Omron Sysmac Studio project 3089-2603A_検査箱詰め装置_CORE_SUB_PIP-02F02NX_20261026D (Sysmac Studio 1.67.0.7, StandardProject)
(* イーサキャット設定完了_20261023I / ST0 供給_20261009A / AutoMode作成_20261008A / IOプログラム作成_20261007B / IOプログラム作成_20261006A / IOプログラム作成_20261005A / IOプログラム作成_20261002A / オリエンタルモータ設定_20261001A / IO設定_20260930A / PLC設定_20260807A *)

# Controller new_Controller_0: NX102-9020 version 1.48
Units and slaves: Node1 : RCGW-ECT(112Byte/112Byte) (E001); Node2 : CVD2A-KED (E002); Node3 : CVD2A-KED (E003); Node5 : RCGW-ECT(112Byte/112Byte) (E005); Node6 : GX-ID1612 (E006); Node7 : GX-ID1612 (E007); Node8 : GX-OD1612 (E008); Node9 : GX-ID1612 (E011); Node10 : GX-OD1612 (E010); ユニット1 : NX-ID6142-6(N1); ユニット2 : NX-ID6142-6(N2); ユニット3 : NX-ID6142-6(N3); ユニット4 : NX-ID6142-6(N4); ユニット5 : NX-ID6142-6(N5); ユニット6 : NX-OD6121-6(N6); ユニット7 : NX-OD6121-6(N7); ユニット8 : NX-OD6121-6(N8)
Axis Stm_A_Rev_Axis000, settings changed from default: AxisType=ServoType, FunctionLimit=SingleAxisPTP, UnitsConversion=EnumElement5, UnitsDenominator=360, MaxVelocity=10000, MaxJogVelocity=10000, HomingMode=BackupAndProximitySignalOn, OriginInputMode=EXT, StartDirection=NegativeDirection, OriginInputDetectionDirection=NegativeDirection, CountMode=EnumElement2, ModuloMAXPosition=360, ModuloMINPosition=0
Axis Stm_A_Rev_Axis001, settings changed from default: AxisNumber=1, AxisType=ServoType, FunctionLimit=SingleAxisPTP, UnitsConversion=EnumElement5, UnitsDenominator=360, MaxVelocity=10000, MaxJogVelocity=10000, HomingMode=BackupAndProximitySignalOn, OriginInputMode=EXT, StartDirection=NegativeDirection, OriginInputDetectionDirection=NegativeDirection, CountMode=EnumElement2, ModuloMAXPosition=360, ModuloMINPosition=0
Axis Stm_B_Rev_Axis002, settings changed from default: AxisNumber=2, AxisType=ServoType, FunctionLimit=SingleAxisPTP, UnitsConversion=EnumElement5, UnitsDenominator=360, MaxVelocity=10000, MaxJogVelocity=10000, HomingMode=BackupAndProximitySignalOn, OriginInputMode=EXT, StartDirection=NegativeDirection, OriginInputDetectionDirection=NegativeDirection, CountMode=EnumElement2, ModuloMAXPosition=360, ModuloMINPosition=0
Axis Stm_B_Rev_Axis003, settings changed from default: AxisNumber=3, AxisType=ServoType, FunctionLimit=SingleAxisPTP, UnitsConversion=EnumElement5, UnitsDenominator=360, MaxVelocity=10000, MaxJogVelocity=10000, HomingMode=BackupAndProximitySignalOn, OriginInputMode=EXT, StartDirection=NegativeDirection, OriginInputDetectionDirection=NegativeDirection, CountMode=EnumElement2, ModuloMAXPosition=360, ModuloMINPosition=0
Task PrimaryTask (priority 4, period or condition 2000): ModeManagement_モード管理, Movements_動作, OtherDevice_外部機器, IO_入出力

TYPE sData : STRUCT
    Dates : STRING[20];  (* 検査日時 *)
    Work_On : BOOL;  (* ワーク有無(0:無 1:有) *)
    Total_Judge : INT;  (* 総合判定(0:無 1:OK 9:NG) *)
    Judgment_Details : INT;  (* NG内容 *)
    HeightData : LREAL;  (* 高さ検査データ *)
END_STRUCT END_TYPE
TYPE ST_RCON_Direct_OUT_Control : STRUCT  (* 出力 制御信号（15BOOL） *)
    Start : BOOL;  (* 開始指令（DSTR/b0・保持10ms以上） *)
    Home : BOOL;  (* 原点復帰指令（HOME/b1） *)
    Pause : BOOL;  (* 一時停止（STP/b2・安全停止ではない） *)
    Reset : BOOL;  (* 異常リセット指令（RES/b3） *)
    ServoOn : BOOL;  (* サーボON指令（SON/b4） *)
    InchingSelect : BOOL;  (* インチング選択（JISL/b5・OFF=ジョグ） *)
    JogSpeedSelect : BOOL;  (* ジョグ速度切替（JVEL/b6） *)
    JogMinus : BOOL;  (* 原点(-)方向ジョグ（JOG-/b7） *)
    JogPlus : BOOL;  (* 反原点方向(+)ジョグ（JOG+/b8） *)
    GainSelect0 : BOOL;  (* ゲイン選択 下位（GSL0/b10） *)
    GainSelect1 : BOOL;  (* ゲイン選択 上位（GSL1/b11） *)
    PushEnable : BOOL;  (* 押付け選択（PUSH/b12・OFF=位置決め） *)
    PushDirection : BOOL;  (* 押付け方向（DIR/b13） *)
    RelativeMove : BOOL;  (* 相対移動選択（INC/b14・OFF=絶対） *)
    BrakeRelease : BOOL;  (* ブレーキ強制解除（BKRL/b15・落下注意） *)
END_STRUCT END_TYPE
TYPE ST_RCON_Direct_IN_Status : STRUCT  (* 入力 状態信号（12BOOL） *)
    PositionDone : BOOL;  (* 位置決め完了（PEND/b0） *)
    HomeDone : BOOL;  (* 原点復帰完了（HEND/b1） *)
    Moving : BOOL;  (* 移動中（MOVE/b2） *)
    Alarm : BOOL;  (* 軸異常（ALM/b3） *)
    ServoReady : BOOL;  (* サーボON状態（SV/b4） *)
    PushMiss : BOOL;  (* 押付け空振り（PSFL/b5） *)
    OverloadWarning : BOOL;  (* 過負荷警告等（ALML/b7） *)
    CommandDone : BOOL;  (* 指令完了（MEND/b8・空振り含む） *)
    Zone1 : BOOL;  (* ゾーン1内（ZONE1/b12） *)
    Zone2 : BOOL;  (* ゾーン2内（ZONE2/b13） *)
    ControllerReady : BOOL;  (* コントローラー準備完了（CRDY/b14） *)
    EmergencyStop : BOOL;  (* 非常停止状態（EMGS/b15・監視用） *)
END_STRUCT END_TYPE
TYPE ST_RCON_Direct_OUT_Axis : STRUCT  (* 1軸分 出力指令（PLC→RCON） *)
    TargetPos_mm : LREAL;  (* 目標位置 [mm] *)
    PositionBand_mm : LREAL;  (* 位置決め幅 [mm] *)
    Speed_mm_s : LREAL;  (* 指令速度 [mm/s] *)
    AccDec_G : LREAL;  (* 共通加減速度 [G] *)
    PushLimit_pct : LREAL;  (* 押付け電流制限 [%] *)
    Control : ST_RCON_Direct_OUT_Control;  (* 出力信号 *)
END_STRUCT END_TYPE
TYPE ST_RCON_Direct_IN_Axis : STRUCT  (* 1軸分 入力情報（RCON→PLC） *)
    ActualPos_mm : LREAL;  (* 現在位置 [mm] *)
    Current_mA : DINT;  (* 指令電流 [mA]（RCON-PC） *)
    ActualSpeed_mm_s : LREAL;  (* 現在速度 [mm/s・符号付き] *)
    AlarmCode : UINT;  (* 軸異常コード *)
    Status : ST_RCON_Direct_IN_Status;  (* 入力信号 *)
    DataValid : BOOL;  (* 入力有効（運転許可とは別） *)
END_STRUCT END_TYPE

VAR_GLOBAL
    In_Sw_EMS1 : BOOL;  (* 【X100】非常停止1(タッチパネル)SW; at IOBus://unit#1/Input Bit 32 bits/Input Bit 00 *)
    In_Sw_EMS2 : BOOL;  (* 【X101】非常停止2(その他)SW; at IOBus://unit#1/Input Bit 32 bits/Input Bit 01 *)
    In_Sw_EMS3 : BOOL;  (* 【X102】非常停止3(その他)SW; at IOBus://unit#1/Input Bit 32 bits/Input Bit 02 *)
    In_Sw_START : BOOL;  (* 【X103】スタートSW; at IOBus://unit#1/Input Bit 32 bits/Input Bit 03 *)
    In_Sw_STOP : BOOL;  (* 【X104】ストップSW; at IOBus://unit#1/Input Bit 32 bits/Input Bit 04 *)
    In_Sw_RESET : BOOL;  (* 【X105】リセットSW; at IOBus://unit#1/Input Bit 32 bits/Input Bit 05 *)
    In_Sen_DOOR_01 : BOOL;  (* 【X108】ドアセンサ1; at IOBus://unit#1/Input Bit 32 bits/Input Bit 08 *)
    In_Sen_DOOR_02 : BOOL;  (* 【X109】ドアセンサ2; at IOBus://unit#1/Input Bit 32 bits/Input Bit 09 *)
    In_Sen_DOOR_03 : BOOL;  (* 【X110】ドアセンサ3; at IOBus://unit#1/Input Bit 32 bits/Input Bit 10 *)
    In_Sen_DOOR_04 : BOOL;  (* 【X111】ドアセンサ4; at IOBus://unit#1/Input Bit 32 bits/Input Bit 11 *)
    In_Sen_DOOR_05 : BOOL;  (* 【X112】ドアセンサ5; at IOBus://unit#1/Input Bit 32 bits/Input Bit 12 *)
    In_Sen_DOOR_06 : BOOL;  (* 【X113】ドアセンサ6; at IOBus://unit#1/Input Bit 32 bits/Input Bit 13 *)
    In_Sen_CV_Alram : BOOL;  (* 【X116】入口 コンベアアラーム; at IOBus://unit#1/Input Bit 32 bits/Input Bit 16 *)
    In_Sen_AIR１_Pressure_01 : BOOL;  (* 【X117】エア圧力(1); at IOBus://unit#1/Input Bit 32 bits/Input Bit 17 *)
    In_Sen_AIR１_Pressure_02 : BOOL;  (* 【X118】エア圧力(2); at IOBus://unit#1/Input Bit 32 bits/Input Bit 18 *)
    In_Sen_AIR１_Pressure_03 : BOOL;  (* 【X119】エア圧力(3); at IOBus://unit#1/Input Bit 32 bits/Input Bit 19 *)
    In_Mtr_Flip_01_A_Error : BOOL;  (* 【X124】A(左側)反転 オリエンタルモータ1 エラー *)
    In_Mtr_Flip_02_A_Error : BOOL;  (* 【X125】A(左側)反転 オリエンタルモータ2 エラー *)
    In_Mtr_Flip_01_B_Error : BOOL;  (* 【X126】B(右側)反転 オリエンタルモータ1 エラー *)
    In_Mtr_Flip_02_B_Error : BOOL;  (* 【X127】B(右側)反転 オリエンタルモータ2 エラー *)
    In_Sen_Accum_CV_B_Full : BOOL;  (* 【X400】B(右側) アキュームCV満; at IOBus://unit#4/Input Bit 32 bits/Input Bit 00 *)
    In_Sen_Accum_CV_A_Arrival : BOOL;  (* 【X201】A(左側) アキューム CV着; at IOBus://unit#2/Input Bit 32 bits/Input Bit 01 *)
    In_Sen_Work_A_Pos_00 : BOOL;  (* 【X202】A(左側)ワーク位置0; at IOBus://unit#2/Input Bit 32 bits/Input Bit 02 *)
    In_Sen_Work_A_Pos_01 : BOOL;  (* 【X203】A(左側)ワーク位置1; at IOBus://unit#2/Input Bit 32 bits/Input Bit 03 *)
    In_Sen_Work_A_Pos_02 : BOOL;  (* 【X204】A(左側)ワーク位置2; at IOBus://unit#2/Input Bit 32 bits/Input Bit 04 *)
    In_Sen_Work_A_Pos_03 : BOOL;  (* 【X205】A(左側)ワーク位置3; at IOBus://unit#2/Input Bit 32 bits/Input Bit 05 *)
    In_Sen_Work_A_Pos_04 : BOOL;  (* 【X206】A(左側)ワーク位置4; at IOBus://unit#2/Input Bit 32 bits/Input Bit 06 *)
    In_Sen_Work_A_Pos_05 : BOOL;  (* 【X207】A(左側)ワーク位置5; at IOBus://unit#2/Input Bit 32 bits/Input Bit 07 *)
    In_Sen_Work_A_Pos_06 : BOOL;  (* 【X208】A(左側)ワーク位置6; at IOBus://unit#2/Input Bit 32 bits/Input Bit 08 *)
    In_Sen_Work_A_Pos_07 : BOOL;  (* 【X209】A(左側)ワーク位置7; at IOBus://unit#2/Input Bit 32 bits/Input Bit 09 *)
    In_Sen_NG1_Tray_01_A_Full : BOOL;  (* 【X210】A(左側) NG1トレイ1満杯; at IOBus://unit#2/Input Bit 32 bits/Input Bit 10 *)
    In_Sen_NG1_Tray_01_A_Full_Warn : BOOL;  (* 【X211】A(左側) NG1トレイ1満杯警告; at IOBus://unit#2/Input Bit 32 bits/Input Bit 11 *)
    In_Sen_NG1_Tray_02_A_Full : BOOL;  (* 【X212】A(左側) NG1トレイ2満杯停止; at IOBus://unit#2/Input Bit 32 bits/Input Bit 12 *)
    In_Sen_NG1_Tray_02_A_Full_Warn : BOOL;  (* 【X213】A(左側) NG1トレイ2満杯警告; at IOBus://unit#2/Input Bit 32 bits/Input Bit 13 *)
    In_Sen_SH_A_Ent : BOOL;  (* 【X214】A(左側) ストックフォルダIN; at IOBus://unit#2/Input Bit 32 bits/Input Bit 14 *)
    In_Sen_SH_A_Ext : BOOL;  (* 【X215】A(左側) ストックフォルダOut; at IOBus://unit#2/Input Bit 32 bits/Input Bit 15 *)
    In_Sen_SH_A_Type_Ent : BOOL;  (* 【X216】A(左側) ストック機種判別IN; at IOBus://unit#2/Input Bit 32 bits/Input Bit 16 *)
    In_Sen_SH_A_Type_Ext : BOOL;  (* 【X217】A(左側) ストック機種判別OUT; at IOBus://unit#2/Input Bit 32 bits/Input Bit 17 *)
    In_SenCY_Sply_Slide_A_H : BOOL;  (* 【X218】A(左側) 供給スライド戻; at IOBus://unit#2/Input Bit 32 bits/Input Bit 18 *)
    In_SenCY_Sply_Slide_A_F : BOOL;  (* 【X219】A(左側) 供給スライド行; at IOBus://unit#2/Input Bit 32 bits/Input Bit 19 *)
    In_SenCY_Sply_Pick_A_H : BOOL;  (* 【X220】A(左側) 供給ピックアップ戻; at IOBus://unit#2/Input Bit 32 bits/Input Bit 20 *)
    In_SenCY_Sply_Pick_A_F : BOOL;  (* 【X221】A(左側) 供給ピックアップ行; at IOBus://unit#2/Input Bit 32 bits/Input Bit 21 *)
    In_SenCY_Sply_Chk_A_H : BOOL;  (* 【X222】A(左側) 供給チャック戻; at IOBus://unit#2/Input Bit 32 bits/Input Bit 22 *)
    In_SenCY_Sply_Chk_A_F : BOOL;  (* 【X223】A(左側) 供給チャック行; at IOBus://unit#2/Input Bit 32 bits/Input Bit 23 *)
    In_SenCY_HgtInsp_Clp_A_H : BOOL;  (* 【X224】A(左側) 高さ検査押え戻; at IOBus://unit#2/Input Bit 32 bits/Input Bit 24 *)
    In_SenCY_HgtInsp_Clp_A_F : BOOL;  (* 【X225】A(左側) 高さ検査押え行; at IOBus://unit#2/Input Bit 32 bits/Input Bit 25 *)
    In_SenCY_HgtInsp_Lf_A_H : BOOL;  (* 【X226】A(左側) 高さ検査持上戻; at IOBus://unit#2/Input Bit 32 bits/Input Bit 26 *)
    In_SenCY_HgtInsp_Lf_A_F : BOOL;  (* 【X227】A(左側) 高さ検査持上行; at IOBus://unit#2/Input Bit 32 bits/Input Bit 27 *)
    In_SenCY_NG1_Pick_A_H : BOOL;  (* 【X228】A(左側) NG1ピックアップ戻; at IOBus://unit#2/Input Bit 32 bits/Input Bit 28 *)
    In_SenCY_NG1_Pick_A_F : BOOL;  (* 【X229】A(左側) NG1ピックアップ行; at IOBus://unit#2/Input Bit 32 bits/Input Bit 29 *)
    In_SenCY_NG1_Chk_A_H : BOOL;  (* 【X230】A(左側) NG1チャック戻; at IOBus://unit#2/Input Bit 32 bits/Input Bit 30 *)
    In_SenCY_NG1_Chk_A_F : BOOL;  (* 【X231】A(左側) NG1チャック行; at IOBus://unit#2/Input Bit 32 bits/Input Bit 31 *)
    In_SenCY_Rev_01_Chk_A_H : BOOL;  (* 【X300】A(左側) 反転1チャック戻; at IOBus://unit#3/Input Bit 32 bits/Input Bit 00 *)
    In_SenCY_Rev_01_Chk_A_F : BOOL;  (* 【X301】A(左側) 反転1チャック行; at IOBus://unit#3/Input Bit 32 bits/Input Bit 01 *)
    In_SenCY_Rev_01_Pick_A_H : BOOL;  (* 【X302】A(左側) 反転1ピックアップ戻; at IOBus://unit#3/Input Bit 32 bits/Input Bit 02 *)
    In_SenCY_Rev_01_Pick_A_F : BOOL;  (* 【X303】A(左側) 反転1ピックアップ行; at IOBus://unit#3/Input Bit 32 bits/Input Bit 03 *)
    In_SenCY_Rev_02_Chk_A_H : BOOL;  (* 【X304】A(左側) 反転2チャック戻; at IOBus://unit#3/Input Bit 32 bits/Input Bit 04 *)
    In_SenCY_Rev_02_Chk_A_F : BOOL;  (* 【X305】A(左側) 反転2チャック行; at IOBus://unit#3/Input Bit 32 bits/Input Bit 05 *)
    In_SenCY_Rev_02_Pick_A_H : BOOL;  (* 【X306】A(左側) 反転2ピックアップ戻; at IOBus://unit#3/Input Bit 32 bits/Input Bit 06 *)
    In_SenCY_Rev_02_Pick_A_F : BOOL;  (* 【X307】A(左側) 反転2ピックアップ行; at IOBus://unit#3/Input Bit 32 bits/Input Bit 07 *)
    In_SenCY_Disc_Chk_A_H : BOOL;  (* 【X308】A(左側) 排出チャック戻; at IOBus://unit#3/Input Bit 32 bits/Input Bit 08 *)
    In_SenCY_Disc_Chk_A_F : BOOL;  (* 【X309】A(左側) 排出チャック行; at IOBus://unit#3/Input Bit 32 bits/Input Bit 09 *)
    In_SenCY_Ejc_SH_Feed_A_H : BOOL;  (* 【X310】A(左側) 排出フォルダ送り戻; at IOBus://unit#3/Input Bit 32 bits/Input Bit 10 *)
    In_SenCY_Ejc_SH_Feed_A_F : BOOL;  (* 【X311】A(左側) 排出フォルダ送り行; at IOBus://unit#3/Input Bit 32 bits/Input Bit 11 *)
    In_SenCY_Pos_01_Stopper_A_H : BOOL;  (* 【X312】A(左側) 位置1ストッパー戻; at IOBus://unit#3/Input Bit 32 bits/Input Bit 12 *)
    In_SenCY_Pos_01_Stopper_A_F : BOOL;  (* 【X313】A(左側) 位置1ストッパー行; at IOBus://unit#3/Input Bit 32 bits/Input Bit 13 *)
    In_SenCY_Pos_02_Stopper_A_H : BOOL;  (* 【X314】A(左側) 位置2ストッパー戻; at IOBus://unit#3/Input Bit 32 bits/Input Bit 14 *)
    In_SenCY_Pos_02_Stopper_A_F : BOOL;  (* 【X315】A(左側) 位置2ストッパー行; at IOBus://unit#3/Input Bit 32 bits/Input Bit 15 *)
    In_SenCY_Pos_03_Stopper_A_H : BOOL;  (* 【X316】A(左側) 位置3ストッパー戻; at IOBus://unit#3/Input Bit 32 bits/Input Bit 16 *)
    In_SenCY_Pos_03_Stopper_A_F : BOOL;  (* 【X317】A(左側) 位置3ストッパー行; at IOBus://unit#3/Input Bit 32 bits/Input Bit 17 *)
    In_SenCY_Pos_04_Stopper_A_H : BOOL;  (* 【X318】A(左側) 位置4ストッパー戻; at IOBus://unit#3/Input Bit 32 bits/Input Bit 18 *)
    In_SenCY_Pos_04_Stopper_A_F : BOOL;  (* 【X319】A(左側) 位置4ストッパー行; at IOBus://unit#3/Input Bit 32 bits/Input Bit 19 *)
    In_SenCY_Pos_05_Stopper_A_H : BOOL;  (* 【X320】A(左側) 位置5ストッパー戻; at IOBus://unit#3/Input Bit 32 bits/Input Bit 20 *)
    In_SenCY_Pos_05_Stopper_A_F : BOOL;  (* 【X321】A(左側) 位置5ストッパー行; at IOBus://unit#3/Input Bit 32 bits/Input Bit 21 *)
    In_SenCY_Pos_06_Stopper_A_H : BOOL;  (* 【X322】A(左側) 位置6ストッパー戻; at IOBus://unit#3/Input Bit 32 bits/Input Bit 22 *)
    In_SenCY_Pos_06_Stopper_A_F : BOOL;  (* 【X323】A(左側) 位置6ストッパー行; at IOBus://unit#3/Input Bit 32 bits/Input Bit 23 *)
    In_SenCY_SH_A_Turn_H : BOOL;  (* 【X324】A(左側) ストックフォルダターン戻; at IOBus://unit#3/Input Bit 32 bits/Input Bit 24 *)
    In_SenCY_SH_A_Turn_F : BOOL;  (* 【X325】A(左側) ストックフォルダターン行; at IOBus://unit#3/Input Bit 32 bits/Input Bit 25 *)
    In_SenCY_NG1_Srt_A_H : BOOL;  (* 【X330】A(左側) NG1仕分け 戻; at IOBus://unit#3/Input Bit 32 bits/Input Bit 30 *)
    In_SenCY_NG1_Srt_A_F : BOOL;  (* 【X331】A(左側) NG1仕分け 行; at IOBus://unit#3/Input Bit 32 bits/Input Bit 31 *)
    In_Sen_Accum_CV_A_Full : BOOL;  (* 【X400】B(右側) アキュームCV満 *)
    In_Sen_Accum_CV_B_Arrival : BOOL;  (* 【X401】B(右側) アキュームCV着; at IOBus://unit#4/Input Bit 32 bits/Input Bit 01 *)
    In_Sen_Work_B_Pos_00 : BOOL;  (* 【X402】B(右側)ワーク位置0; at IOBus://unit#4/Input Bit 32 bits/Input Bit 02 *)
    In_Sen_Work_B_Pos_01 : BOOL;  (* 【X403】B(右側)ワーク位置1; at IOBus://unit#4/Input Bit 32 bits/Input Bit 03 *)
    In_Sen_Work_B_Pos_02 : BOOL;  (* 【X404】B(右側)ワーク位置2; at IOBus://unit#4/Input Bit 32 bits/Input Bit 04 *)
    In_Sen_Work_B_Pos_03 : BOOL;  (* 【X405】B(右側)ワーク位置3; at IOBus://unit#4/Input Bit 32 bits/Input Bit 05 *)
    In_Sen_Work_B_Pos_04 : BOOL;  (* 【X406】B(右側)ワーク位置4; at IOBus://unit#4/Input Bit 32 bits/Input Bit 06 *)
    In_Sen_Work_B_Pos_05 : BOOL;  (* 【X407】B(右側)ワーク位置5; at IOBus://unit#4/Input Bit 32 bits/Input Bit 07 *)
    In_Sen_Work_B_Pos_06 : BOOL;  (* 【X408】B(右側)ワーク位置6; at IOBus://unit#4/Input Bit 32 bits/Input Bit 08 *)
    In_Sen_Work_B_Pos_07 : BOOL;  (* 【X409】B(右側)ワーク位置7; at IOBus://unit#4/Input Bit 32 bits/Input Bit 09 *)
    In_Sen_NG1_Tray_01_B_Full : BOOL;  (* 【X410】B(右側) NG1トレイ1満杯; at IOBus://unit#4/Input Bit 32 bits/Input Bit 10 *)
    In_Sen_NG1_Tray_01_B_Full_Warn : BOOL;  (* 【X411】B(右側) NG1トレイ1満杯警告; at IOBus://unit#4/Input Bit 32 bits/Input Bit 11 *)
    In_Sen_NG1_Tray_02_B_Full : BOOL;  (* 【X412】B(右側) NG1トレイ2満杯停止; at IOBus://unit#4/Input Bit 32 bits/Input Bit 12 *)
    In_Sen_NG1_Tray_02_B_Full_Warn : BOOL;  (* 【X413】B(右側) NG1トレイ2満杯警告; at IOBus://unit#4/Input Bit 32 bits/Input Bit 13 *)
    In_Sen_SH_B_Ent : BOOL;  (* 【X414】B(右側) ストックフォルダIN; at IOBus://unit#4/Input Bit 32 bits/Input Bit 14 *)
    In_Sen_SH_B_Ext : BOOL;  (* 【X415】B(右側) ストックフォルダOut; at IOBus://unit#4/Input Bit 32 bits/Input Bit 15 *)
    In_Sen_SH_B_Type_Ent : BOOL;  (* 【X416】B(右側) ストック機種判別IN; at IOBus://unit#4/Input Bit 32 bits/Input Bit 16 *)
    In_Sen_SH_B_Type_Ext : BOOL;  (* 【X417】B(右側) ストック機種判別OUT; at IOBus://unit#4/Input Bit 32 bits/Input Bit 17 *)
    In_SenCY_Sply_Slide_B_H : BOOL;  (* 【X418】B(右側) 供給スライド戻; at IOBus://unit#4/Input Bit 32 bits/Input Bit 18 *)
    In_SenCY_Sply_Slide_B_F : BOOL;  (* 【X419】B(右側) 供給スライド行; at IOBus://unit#4/Input Bit 32 bits/Input Bit 19 *)
    In_SenCY_Sply_Pick_B_H : BOOL;  (* 【X420】B(右側) 供給ピックアップ戻; at IOBus://unit#4/Input Bit 32 bits/Input Bit 20 *)
    In_SenCY_Sply_Pick_B_F : BOOL;  (* 【X421】B(右側) 供給ピックアップ行; at IOBus://unit#4/Input Bit 32 bits/Input Bit 21 *)
    In_SenCY_Sply_Chk_B_H : BOOL;  (* 【X422】B(右側) 供給チャック閉 戻; at IOBus://unit#4/Input Bit 32 bits/Input Bit 22 *)
    In_SenCY_Sply_Chk_B_F : BOOL;  (* 【X423】B(右側) 供給チャック開 行; at IOBus://unit#4/Input Bit 32 bits/Input Bit 23 *)
    In_SenCY_HgtInsp_Clp_B_H : BOOL;  (* 【X424】B(右側) 高さ検査押え戻; at IOBus://unit#4/Input Bit 32 bits/Input Bit 24 *)
    In_SenCY_HgtInsp_Clp_B_F : BOOL;  (* 【X425】B(右側) 高さ検査押え行; at IOBus://unit#4/Input Bit 32 bits/Input Bit 25 *)
    In_SenCY_HgtInsp_Lf_B_H : BOOL;  (* 【X426】B(右側) 高さ検査持上戻; at IOBus://unit#4/Input Bit 32 bits/Input Bit 26 *)
    In_SenCY_HgtInsp_Lf_B_F : BOOL;  (* 【X427】B(右側) 高さ検査持上行; at IOBus://unit#4/Input Bit 32 bits/Input Bit 27 *)
    In_SenCY_NG1_Pick_B_H : BOOL;  (* 【X428】B(右側) NG1ピックアップ戻; at IOBus://unit#4/Input Bit 32 bits/Input Bit 28 *)
    In_SenCY_NG1_Pick_B_F : BOOL;  (* 【X429】B(右側) NG1ピックアップ行; at IOBus://unit#4/Input Bit 32 bits/Input Bit 29 *)
    In_SenCY_NG1_Chk_B_H : BOOL;  (* 【X430】B(右側) NG1チャック閉 戻; at IOBus://unit#4/Input Bit 32 bits/Input Bit 30 *)
    In_SenCY_NG1_Chk_B_F : BOOL;  (* 【X431】B(右側) NG1チャック開 行; at IOBus://unit#4/Input Bit 32 bits/Input Bit 31 *)
    In_SenCY_Rev_01_Chk_B_H : BOOL;  (* 【X500】B(右側)ST4 反転1チャック閉 戻; at IOBus://unit#5/Input Bit 32 bits/Input Bit 00 *)
    In_SenCY_Rev_01_Chk_B_F : BOOL;  (* 【X501】B(右側)ST4 反転1チャック開 行; at IOBus://unit#5/Input Bit 32 bits/Input Bit 01 *)
    In_SenCY_Rev_01_Pick_B_H : BOOL;  (* 【X502】B(右側)ST4 反転1ピックアップ戻; at IOBus://unit#5/Input Bit 32 bits/Input Bit 02 *)
    In_SenCY_Rev_01_Pick_B_F : BOOL;  (* 【X503】B(右側)ST4 反転1ピックアップ行; at IOBus://unit#5/Input Bit 32 bits/Input Bit 03 *)
    In_SenCY_Rev_02_Chk_B_H : BOOL;  (* 【X504】B(右側)ST6 反転2チャック閉 戻; at IOBus://unit#5/Input Bit 32 bits/Input Bit 04 *)
    In_SenCY_Rev_02_Chk_B_F : BOOL;  (* 【X505】B(右側)ST6 反転2チャック開 行; at IOBus://unit#5/Input Bit 32 bits/Input Bit 05 *)
    In_SenCY_Rev_02_Pick_B_H : BOOL;  (* 【X506】B(右側)ST6 反転2ピックアップ戻; at IOBus://unit#5/Input Bit 32 bits/Input Bit 06 *)
    In_SenCY_Rev_02_Pick_B_F : BOOL;  (* 【X507】B(右側)ST6 反転2ピックアップ行; at IOBus://unit#5/Input Bit 32 bits/Input Bit 07 *)
    In_SenCY_Disc_Chk_B_H : BOOL;  (* 【X508】B(右側) 排出チャック閉 戻; at IOBus://unit#5/Input Bit 32 bits/Input Bit 08 *)
    In_SenCY_Disc_Chk_B_F : BOOL;  (* 【X509】B(右側) 排出チャック開 行; at IOBus://unit#5/Input Bit 32 bits/Input Bit 09 *)
    In_SenCY_Ejc_SH_Feed_B_F : BOOL;  (* 【X510】B(右側) 排出フォルダ送り戻; at IOBus://unit#5/Input Bit 32 bits/Input Bit 10 *)
    In_SenCY_Ejc_SH_Feed_B_H : BOOL;  (* 【X511】B(右側) 排出フォルダ送り行; at IOBus://unit#5/Input Bit 32 bits/Input Bit 11 *)
    In_SenCY_Pos_01_Stopper_B_H : BOOL;  (* 【X512】B(右側) 位置1ストッパー戻; at IOBus://unit#5/Input Bit 32 bits/Input Bit 12 *)
    In_SenCY_Pos_01_Stopper_B_F : BOOL;  (* 【X513】B(右側) 位置1ストッパー行; at IOBus://unit#5/Input Bit 32 bits/Input Bit 13 *)
    In_SenCY_Pos_02_Stopper_B_H : BOOL;  (* 【X514】B(右側) 位置2ストッパー戻; at IOBus://unit#5/Input Bit 32 bits/Input Bit 14 *)
    In_SenCY_Pos_02_Stopper_B_F : BOOL;  (* 【X515】B(右側) 位置2ストッパー行; at IOBus://unit#5/Input Bit 32 bits/Input Bit 15 *)
    In_SenCY_Pos_03_Stopper_B_H : BOOL;  (* 【X516】B(右側) 位置3ストッパー戻; at IOBus://unit#5/Input Bit 32 bits/Input Bit 16 *)
    In_SenCY_Pos_03_Stopper_B_F : BOOL;  (* 【X517】B(右側) 位置3ストッパー行; at IOBus://unit#5/Input Bit 32 bits/Input Bit 17 *)
    In_SenCY_Pos_04_Stopper_B_H : BOOL;  (* 【X518】B(右側) 位置4ストッパー戻; at IOBus://unit#5/Input Bit 32 bits/Input Bit 18 *)
    In_SenCY_Pos_04_Stopper_B_F : BOOL;  (* 【X519】B(右側) 位置4ストッパー行; at IOBus://unit#5/Input Bit 32 bits/Input Bit 19 *)
    In_SenCY_Pos_05_Stopper_B_H : BOOL;  (* 【X520】B(右側) 位置5ストッパー戻; at IOBus://unit#5/Input Bit 32 bits/Input Bit 20 *)
    In_SenCY_Pos_05_Stopper_B_F : BOOL;  (* 【X521】B(右側) 位置5ストッパー行; at IOBus://unit#5/Input Bit 32 bits/Input Bit 21 *)
    In_SenCY_Pos_06_Stopper_B_H : BOOL;  (* 【X522】B(右側) 位置6ストッパー戻; at IOBus://unit#5/Input Bit 32 bits/Input Bit 22 *)
    In_SenCY_Pos_06_Stopper_B_F : BOOL;  (* 【X523】B(右側) 位置6ストッパー行; at IOBus://unit#5/Input Bit 32 bits/Input Bit 23 *)
    In_SenCY_SH_B_Turn_H : BOOL;  (* 【X524】B(右側) ストックフォルダターン戻; at IOBus://unit#5/Input Bit 32 bits/Input Bit 24 *)
    In_SenCY_SH_B_Turn_F : BOOL;  (* 【X525】B(右側) ストックフォルダターン行; at IOBus://unit#5/Input Bit 32 bits/Input Bit 25 *)
    In_SenCY_NG1_Srt_B_H : BOOL;  (* 【X530】B(右側) NG1 仕分け 戻; at IOBus://unit#5/Input Bit 32 bits/Input Bit 30 *)
    In_SenCY_NG1_Srt_B_F : BOOL;  (* 【X531】B(右側) NG1 仕分け 行; at IOBus://unit#5/Input Bit 32 bits/Input Bit 31 *)
    In_Sen_Supply_Container_Exist : BOOL;  (* 【X1000】供給部コンテナ有; at ECAT://node#6/Read input 1st word/In Bit00 *)
    In_Sen_Destacker_Stage_01_Exist : BOOL;  (* 【X1001】段バラシ1段目有; at ECAT://node#6/Read input 1st word/In Bit01 *)
    In_Sen_Destacker_Stage_02_Exist : BOOL;  (* 【X1002】段バラシ2段目有; at ECAT://node#6/Read input 1st word/In Bit02 *)
    In_Sen_Container_Arrival : BOOL;  (* 【X1003】コンテナ到着; at ECAT://node#6/Read input 1st word/In Bit03 *)
    In_Sen_Container_Direction_Check : BOOL;  (* 【X1004】コンテナ方向確認; at ECAT://node#6/Read input 1st word/In Bit04 *)
    In_Sen_Container_Pass : BOOL;  (* 【X1005】コンテナ通過; at ECAT://node#6/Read input 1st word/In Bit05 *)
    In_Sen_Container_Full : BOOL;  (* 【X1006】コンテナ満杯; at ECAT://node#6/Read input 1st word/In Bit06 *)
    In_Sen_Tray_Direction_Check : BOOL;  (* 【X1007】コンテナトレイ方向; at ECAT://node#6/Read input 1st word/In Bit07 *)
    In_SenCY_Empty_Container_CY_H : BOOL;  (* 【X1010】空コンテナ送り 戻; at ECAT://node#6/Read input 1st word/In Bit10 *)
    In_SenCY_Empty_Container_CY_F : BOOL;  (* 【X1011】空コンテナ送り 行; at ECAT://node#6/Read input 1st word/In Bit11 *)
    In_SenCY_Sep_Claw1_H : BOOL;  (* 【X1012】段バラシ爪1 戻; at ECAT://node#6/Read input 1st word/In Bit12 *)
    In_SenCY_Sep_Claw1_F : BOOL;  (* 【X1013】段バラシ爪1 行; at ECAT://node#6/Read input 1st word/In Bit13 *)
    In_SenCY_Sep_Claw2_H : BOOL;  (* 【X1014】段バラシ爪2 戻; at ECAT://node#6/Read input 1st word/In Bit14 *)
    In_SenCY_Sep_Claw2_F : BOOL;  (* 【X1015】段バラシ爪2 行; at ECAT://node#6/Read input 1st word/In Bit15 *)
    In_SenCY_Ejc_Cont1_H : BOOL;  (* 【X1016】コンテナ排出1 戻; at ECAT://node#7/Read input 1st word/In Bit00 *)
    In_SenCY_Ejc_Cont1_F : BOOL;  (* 【X1017】コンテナ排出1 行; at ECAT://node#7/Read input 1st word/In Bit01 *)
    In_SenCY_Ejc_Cont2_H : BOOL;  (* 【X1018】コンテナ排出2 戻; at ECAT://node#7/Read input 1st word/In Bit02 *)
    In_SenCY_Ejc_Cont2_F : BOOL;  (* 【X1019】コンテナ排出2 行; at ECAT://node#7/Read input 1st word/In Bit03 *)
    In_SenCY_Box_Chk_H : BOOL;  (* 【X1020】箱入れチャック 戻; at ECAT://node#7/Read input 1st word/In Bit04 *)
    In_SenCY_Box_Chk_F : BOOL;  (* 【X1021】箱入れチャック 行; at ECAT://node#7/Read input 1st word/In Bit05 *)
    In_SenCY_Srt_Stopper_H : BOOL;  (* 【X1022】コンテナ仕分けストッパー 戻; at ECAT://node#7/Read input 1st word/In Bit06 *)
    In_SenCY_Srt_Stopper_F : BOOL;  (* 【X1023】コンテナ仕分けストッパー 行; at ECAT://node#7/Read input 1st word/In Bit07 *)
    In_SenCY_Srt_Feed_H : BOOL;  (* 【X1024】コンテナ仕分け送り 戻; at ECAT://node#7/Read input 1st word/In Bit08 *)
    In_SenCY_Srt_Feed_F : BOOL;  (* 【X1025】コンテナ仕分け送り 行; at ECAT://node#7/Read input 1st word/In Bit09 *)
    Out_CYw_Hnd_Feed_A_H : BOOL;  (* 【Y1300】A(左側) コンベア受渡送り戻; at ECAT://node#10/Write output 1st word/Out Bit00 *)
    Out_CYw_Hnd_Feed_A_F : BOOL;  (* 【Y1301】A(左側) コンベア受渡送り行; at ECAT://node#10/Write output 1st word/Out Bit01 *)
    Out_CYw_Hnd_Feed_B_H : BOOL;  (* 【Y1302】B(右側) コンベア受渡送り戻; at ECAT://node#10/Write output 1st word/Out Bit02 *)
    Out_CYw_Hnd_Feed_B_F : BOOL;  (* 【Y1303】B(右側) コンベア受渡送り行; at ECAT://node#10/Write output 1st word/Out Bit03 *)
    In_Sen_Unl_Conv_A_Pass : BOOL;  (* 【X1100】A(左側) 取出しコンベア 通過; at ECAT://node#9/Read input 1st word/In Bit00 *)
    In_Sen_Unl_Conv_B_Pass : BOOL;  (* 【X1101】B(右側) 取出しコンベア 通過; at ECAT://node#9/Read input 1st word/In Bit01 *)
    In_Sen_Trs_Conv_A_Arrival : BOOL;  (* 【X1102】A(左側) 搬送コンベア到着; at ECAT://node#9/Read input 1st word/In Bit02 *)
    In_Sen_Trs_Conv_B_Arrival : BOOL;  (* 【X1103】B(右側) 搬送コンベア到着; at ECAT://node#9/Read input 1st word/In Bit03 *)
    In_SenCY_Hnd_Feed_A_H : BOOL;  (* 【X1104】A(左側) コンベア受渡送り戻; at ECAT://node#9/Read input 1st word/In Bit04 *)
    In_SenCY_Hnd_Feed_A_F : BOOL;  (* 【X1105】A(左側) コンベア受渡送り行; at ECAT://node#9/Read input 1st word/In Bit05 *)
    In_SenCY_Hnd_Feed_B_H : BOOL;  (* 【X1106】B(右側) コンベア受渡送り戻; at ECAT://node#9/Read input 1st word/In Bit06 *)
    In_SenCY_Hnd_Feed_B_F : BOOL;  (* 【X1107】B(右側) コンベア受渡送り行; at ECAT://node#9/Read input 1st word/In Bit07 *)
    Out_CYw_Empty_Container_CY_H : BOOL;  (* 【Y1200】空コンテナ送り 戻; at ECAT://node#8/Write output 1st word/Out Bit00 *)
    Out_CYw_Empty_Container_CY_F : BOOL;  (* 【Y1201】空コンテナ送り 行; at ECAT://node#8/Write output 1st word/Out Bit01 *)
    Out_CYw_Sep_Claw_F : BOOL;  (* 【Y1203】段バラシ爪 行; at ECAT://node#8/Write output 1st word/Out Bit03 *)
    Out_CYw_Sep_Claw_H : BOOL;  (* 【Y1202】段バラシ爪 戻; at ECAT://node#8/Write output 1st word/Out Bit02 *)
    Out_CYw_Ejc_Cont_H : BOOL;  (* 【Y1204】コンテナ排出 戻; at ECAT://node#8/Write output 1st word/Out Bit04 *)
    Out_CYw_Ejc_Cont_F : BOOL;  (* 【Y1205】コンテナ排出 行; at ECAT://node#8/Write output 1st word/Out Bit05 *)
    Out_CYw_Box_Chuck_H : BOOL;  (* 【Y1206】箱入れチャック 戻; at ECAT://node#8/Write output 1st word/Out Bit06 *)
    Out_CYw_Box_Chuck_F : BOOL;  (* 【Y1207】箱入れチャック 行; at ECAT://node#8/Write output 1st word/Out Bit07 *)
    Out_CYw_Srt_Stopper_H : BOOL;  (* 【Y1208】コンテナ仕分けストッパー 戻; at ECAT://node#8/Write output 1st word/Out Bit08 *)
    Out_CYw_Srt_Stopper_F : BOOL;  (* 【Y1209】コンテナ仕分けストッパー 行; at ECAT://node#8/Write output 1st word/Out Bit09 *)
    Out_CYw_Srt_Feed_H : BOOL;  (* 【Y1210】コンテナ仕分け送り 戻; at ECAT://node#8/Write output 1st word/Out Bit10 *)
    Out_CYw_Srt_Feed_F : BOOL;  (* 【Y1211】コンテナ仕分け送り 行; at ECAT://node#8/Write output 1st word/Out Bit11 *)
    E002_Axis1_Receive_PDO_mapping_1_Controlword_6040_00 : UINT;
    E002_Axis1_Receive_PDO_mapping_1_Target_position_607A_00 : DINT;
    E002_Axis1_Receive_PDO_mapping_1_Modes_of_operation_6060_00 : SINT;
    E002_Axis1_Receive_PDO_mapping_1_Profile_velocity_6081_00 : UDINT;
    E002_Axis2_Receive_PDO_mapping_1_Controlword_6840_00 : UINT;
    E002_Axis2_Receive_PDO_mapping_1_Target_position_687A_00 : DINT;
    E002_Axis2_Receive_PDO_mapping_1_Modes_of_operation_6860_00 : SINT;
    E002_Axis2_Receive_PDO_mapping_1_Profile_velocity_6881_00 : UDINT;
    E002_Axis1_Transmit_PDO_mapping_Statusword_6041_00 : UINT;
    E002_Axis1_Transmit_PDO_mapping_Position_actual_value_6064_00 : DINT;
    E002_Axis1_Transmit_PDO_mapping_Modes_of_operation_display_6061_00 : SINT;
    E002_Axis2_Transmit_PDO_mapping_Statusword_6841_00 : UINT;
    E002_Axis2_Transmit_PDO_mapping_Position_actual_value_6864_00 : DINT;
    E002_Axis2_Transmit_PDO_mapping_Modes_of_operation_display_6861_00 : SINT;
    E003_Axis1_Receive_PDO_mapping_1_Controlword_6040_00 : UINT;
    E003_Axis1_Receive_PDO_mapping_1_Target_position_607A_00 : DINT;
    E003_Axis1_Receive_PDO_mapping_1_Modes_of_operation_6060_00 : SINT;
    E003_Axis1_Receive_PDO_mapping_1_Profile_velocity_6081_00 : UDINT;
    E003_Axis2_Receive_PDO_mapping_1_Controlword_6840_00 : UINT;
    E003_Axis2_Receive_PDO_mapping_1_Target_position_687A_00 : DINT;
    E003_Axis2_Receive_PDO_mapping_1_Modes_of_operation_6860_00 : SINT;
    E003_Axis2_Receive_PDO_mapping_1_Profile_velocity_6881_00 : UDINT;
    E003_Axis1_Transmit_PDO_mapping_Statusword_6041_00 : UINT;
    E003_Axis1_Transmit_PDO_mapping_Position_actual_value_6064_00 : DINT;
    E003_Axis1_Transmit_PDO_mapping_Modes_of_operation_display_6061_00 : SINT;
    E003_Axis2_Transmit_PDO_mapping_Statusword_6841_00 : UINT;
    E003_Axis2_Transmit_PDO_mapping_Position_actual_value_6864_00 : DINT;
    E003_Axis2_Transmit_PDO_mapping_Modes_of_operation_display_6861_00 : SINT;
END_VAR
VAR_GLOBAL CONSTANT
    Stm_A_Rev_Axis000 : _sAXIS_REF;  (* at MC://_MC_AX[0] *)
    Stm_A_Rev_Axis001 : _sAXIS_REF;  (* at MC://_MC_AX[1] *)
END_VAR
VAR_GLOBAL
    Out_SW_Start_LP_GREEN : BOOL;  (* 【Y600】SWスタートランプ緑; at IOBus://unit#6/Output Bit 32 bits/Output Bit 00 *)
    Out_SW_Stop_LP_RED : BOOL;  (* 【Y601】SWストップランプ赤; at IOBus://unit#6/Output Bit 32 bits/Output Bit 01 *)
    Out_SW_Reset_LP_Orange : BOOL;  (* 【Y602】SW リセットランプ橙; at IOBus://unit#6/Output Bit 32 bits/Output Bit 02 *)
    Out_Sg_LP_GREEN : BOOL;  (* 【Y603】シグナルタワー緑; at IOBus://unit#6/Output Bit 32 bits/Output Bit 03 *)
    Out_Sg_LP_RED : BOOL;  (* 【Y604】シグナルタワー赤; at IOBus://unit#6/Output Bit 32 bits/Output Bit 04 *)
    Out_Sg_LP_ORANGE : BOOL;  (* 【Y605】シグナルタワー橙; at IOBus://unit#6/Output Bit 32 bits/Output Bit 05 *)
    Out_Sg_BUZZER : BOOL;  (* 【Y606】シグナルタワーブザー; at IOBus://unit#6/Output Bit 32 bits/Output Bit 06 *)
    Out_Acc_Conv_Run : BOOL;  (* 【Y607】アキューム コンベア運転ON; at IOBus://unit#6/Output Bit 32 bits/Output Bit 07 *)
    Out_Accum_Cv_PowerOn : BOOL;  (* 【Y609】アキューム コンベア電源ON *)
    Out_Insp_Cv_A_Run : BOOL;  (* 【Y610】A(左側) 検査コンベア運転ON; at IOBus://unit#6/Output Bit 32 bits/Output Bit 10 *)
    Out_Insp_Cv_A_RESET : BOOL;  (* 【Y611】A(左側) 検査コンベア リセット *)
    Out_Insp_Cv_A_PowerOn : BOOL;  (* 【Y612】A(左側) 検査コンベア 電源ON *)
    Out_Insp_Cv_B_Run : BOOL;  (* 【Y613】B(右側) 検査コンベア運転ON; at IOBus://unit#6/Output Bit 32 bits/Output Bit 13 *)
    Out_Insp_Cv_B_RESET : BOOL;  (* 【Y614】B(右側) 検査コンベア リセット *)
    Out_Insp_Cv_B_PowerOn : BOOL;  (* 【Y615】B(右側) 検査コンベア 電源ON *)
    Out_Accum_Cv_RESET : BOOL;  (* 【Y608】アキューム コンベア リセット *)
    Out_CYw_Sply_Slide_A_H : BOOL;  (* 【Y616】A(左側) 供給スライド戻; at IOBus://unit#6/Output Bit 32 bits/Output Bit 16 *)
    Out_CYw_Sply_Slide_A_F : BOOL;  (* 【Y617】A(左側) 供給スライド行; at IOBus://unit#6/Output Bit 32 bits/Output Bit 17 *)
    Out_CYw_Sply_Pick_A_H : BOOL;  (* 【Y618】A(左側) 供給ピックアップ戻; at IOBus://unit#6/Output Bit 32 bits/Output Bit 18 *)
    Out_CYw_Sply_Pick_A_F : BOOL;  (* 【Y619】A(左側) 供給ピックアップ行; at IOBus://unit#6/Output Bit 32 bits/Output Bit 19 *)
    Out_CYw_Sup_Chuck_A_Cl_H : BOOL;  (* 【Y620】A(左側) 供給チャック閉 戻; at IOBus://unit#6/Output Bit 32 bits/Output Bit 20 *)
    Out_CYw_Sup_Chuck_A_Op_F : BOOL;  (* 【Y621】A(左側) 供給チャック開 行; at IOBus://unit#6/Output Bit 32 bits/Output Bit 21 *)
    Out_CYw_Sply_Slide_B_H : BOOL;  (* 【Y622】B(右側) 供給スライド戻; at IOBus://unit#6/Output Bit 32 bits/Output Bit 22 *)
    Out_CYw_Sply_Slide_B_F : BOOL;  (* 【Y623】B(右側) 供給スライド行; at IOBus://unit#6/Output Bit 32 bits/Output Bit 23 *)
    Out_CYw_Sply_Pick_B_H : BOOL;  (* 【Y624】B(右側) 供給ピックアップ戻; at IOBus://unit#6/Output Bit 32 bits/Output Bit 24 *)
    Out_CYw_Sply_Pick_B_F : BOOL;  (* 【Y625】B(右側) 供給ピックアップ行; at IOBus://unit#6/Output Bit 32 bits/Output Bit 25 *)
    Out_CYw_Sup_Chuck_B_Cl_H : BOOL;  (* 【Y626】B(右側) 供給チャック閉 戻; at IOBus://unit#6/Output Bit 32 bits/Output Bit 26 *)
    Out_CYw_Sup_Chuck_B_Op_F : BOOL;  (* 【Y627】B(右側) 供給チャック開 行; at IOBus://unit#6/Output Bit 32 bits/Output Bit 27 *)
    Out_CYw_HgtInsp_Clp_A_H : BOOL;  (* 【Y700】A(左側) 高さ検査押え戻; at IOBus://unit#7/Output Bit 32 bits/Output Bit 00 *)
    Out_CYw_HgtInsp_Clp_A_F : BOOL;  (* 【Y701】A(左側) 高さ検査押え行; at IOBus://unit#7/Output Bit 32 bits/Output Bit 01 *)
    Out_CYw_HgtInsp_Lf_A_H : BOOL;  (* 【Y702】A(左側) 高さ検査持上戻; at IOBus://unit#7/Output Bit 32 bits/Output Bit 02 *)
    Out_CYw_HgtInsp_Lf_A_F : BOOL;  (* 【Y703】A(左側) 高さ検査持上行; at IOBus://unit#7/Output Bit 32 bits/Output Bit 03 *)
    Out_CYw_NG1_Pick_A_H : BOOL;  (* 【Y704】A(左側) NG1ピックアップ戻; at IOBus://unit#7/Output Bit 32 bits/Output Bit 04 *)
    Out_CYw_NG1_Pick_A_F : BOOL;  (* 【Y705】A(左側) NG1ピックアップ 行; at IOBus://unit#7/Output Bit 32 bits/Output Bit 05 *)
    Out_CYw_NG1_Chk_A_H : BOOL;  (* 【Y706】A(左側) NG1チャック戻; at IOBus://unit#7/Output Bit 32 bits/Output Bit 06 *)
    Out_CYw_NG1_Chk_A_F : BOOL;  (* 【Y707】A(左側) NG1チャック行; at IOBus://unit#7/Output Bit 32 bits/Output Bit 07 *)
    Out_CYw_Rev_01_Chk_A_H : BOOL;  (* 【Y708】A(左側)ST4 反転1チャック閉; at IOBus://unit#7/Output Bit 32 bits/Output Bit 08 *)
    Out_CYw_Rev_01_Chk_A_F : BOOL;  (* 【Y709】A(左側)ST4 反転1チャック開; at IOBus://unit#7/Output Bit 32 bits/Output Bit 09 *)
    Out_CYw_Rev_01_Pick_A_H : BOOL;  (* 【Y710】A(左側)ST4 反転1ピックアップ戻; at IOBus://unit#7/Output Bit 32 bits/Output Bit 10 *)
    Out_CYw_Rev_01_Pick_A_F : BOOL;  (* 【Y711】A(左側)ST4 反転1ピックアップ行; at IOBus://unit#7/Output Bit 32 bits/Output Bit 11 *)
    Out_CYw_Rev_02_Chk_A_H : BOOL;  (* 【Y712】A(左側)ST6 反転2チャック閉 戻; at IOBus://unit#7/Output Bit 32 bits/Output Bit 12 *)
    Out_CYw_Rev_02_Chk_A_F : BOOL;  (* 【Y713】A(左側)ST6 反転2チャック開 行; at IOBus://unit#7/Output Bit 32 bits/Output Bit 13 *)
    Out_CYw_Rev_02_Pick_A_H : BOOL;  (* 【Y714】A(左側)ST6 反転2ピックアップ戻; at IOBus://unit#7/Output Bit 32 bits/Output Bit 14 *)
    Out_CYw_Rev_02_Pick_A_F : BOOL;  (* 【Y715】A(左側)ST6 反転2ピックアップ行; at IOBus://unit#7/Output Bit 32 bits/Output Bit 15 *)
    Out_CYw_Disc_Chk_A_H : BOOL;  (* 【Y716】A(左側) 排出チャック閉 戻; at IOBus://unit#7/Output Bit 32 bits/Output Bit 16 *)
    Out_CYw_Disc_Chk_A_F : BOOL;  (* 【Y717】A(左側) 排出チャック開 行; at IOBus://unit#7/Output Bit 32 bits/Output Bit 17 *)
    Out_CYw_Ejc_Hldr_Feed_A_F : BOOL;  (* 【Y719】A(左側) 排出フォルダ送り行; at IOBus://unit#7/Output Bit 32 bits/Output Bit 19 *)
    Out_CYw_Ejc_Hldr_Feed_A_H : BOOL;  (* 【Y718】A(左側) 排出フォルダ送り戻; at IOBus://unit#7/Output Bit 32 bits/Output Bit 18 *)
    Out_CYS_Pos_01_Stopper_A : BOOL;  (* 【Y720】A(左側) 位置1ストッパー; at IOBus://unit#7/Output Bit 32 bits/Output Bit 20 *)
    Out_CYS_Pos_02_Stopper_A : BOOL;  (* 【Y721】A(左側) 位置2ストッパー; at IOBus://unit#7/Output Bit 32 bits/Output Bit 21 *)
    Out_CYS_Pos_03_Stopper_A : BOOL;  (* 【Y722】A(左側) 位置3ストッパー; at IOBus://unit#7/Output Bit 32 bits/Output Bit 22 *)
    Out_CYS_Pos_04_Stopper_A : BOOL;  (* 【Y723】A(左側) 位置4ストッパー; at IOBus://unit#7/Output Bit 32 bits/Output Bit 23 *)
    Out_CYS_Pos_05_Stopper_A : BOOL;  (* 【Y724】A(左側) 位置5ストッパー; at IOBus://unit#7/Output Bit 32 bits/Output Bit 24 *)
    Out_CYS_Pos_06_Stopper_A : BOOL;  (* 【Y725】A(左側) 位置6ストッパー; at IOBus://unit#7/Output Bit 32 bits/Output Bit 25 *)
    Out_CYw_SH_A_Turn_H : BOOL;  (* 【Y726】A(左側) ストックフォルダターン戻; at IOBus://unit#7/Output Bit 32 bits/Output Bit 26 *)
    Out_CYw_SH_A_Turn_F : BOOL;  (* 【Y727】A(左側) ストックフォルダターン行; at IOBus://unit#7/Output Bit 32 bits/Output Bit 27 *)
    Out_CYw_NG1_Srt_A_H : BOOL;  (* 【Y728】A(左側) NG1仕分け 戻; at IOBus://unit#7/Output Bit 32 bits/Output Bit 28 *)
    Out_CYw_NG1_Srt_A_F : BOOL;  (* 【Y729】A(左側) NG1仕分け 行; at IOBus://unit#7/Output Bit 32 bits/Output Bit 29 *)
    Out_CYw_HgtInsp_Clp_B_H : BOOL;  (* 【Y800】B(右側) 高さ検査押え戻; at IOBus://unit#8/Output Bit 32 bits/Output Bit 00 *)
    Out_CYw_HgtInsp_Clp_B_F : BOOL;  (* 【Y801】B(右側) 高さ検査押え行; at IOBus://unit#8/Output Bit 32 bits/Output Bit 01 *)
    Out_CYw_HgtInsp_Lf_B_H : BOOL;  (* 【Y802】B(右側) 高さ検査持上戻; at IOBus://unit#8/Output Bit 32 bits/Output Bit 02 *)
    Out_CYw_HgtInsp_Lf_B_F : BOOL;  (* 【Y803】B(右側) 高さ検査持上行; at IOBus://unit#8/Output Bit 32 bits/Output Bit 03 *)
    Out_CYw_NG1_Pick_B_H : BOOL;  (* 【Y804】B(右側) NG1ピックアップ戻; at IOBus://unit#8/Output Bit 32 bits/Output Bit 04 *)
    Out_CYw_NG1_Pick_B_F : BOOL;  (* 【Y805】B(右側) NG1ピックアップ行; at IOBus://unit#8/Output Bit 32 bits/Output Bit 05 *)
    Out_CYw_NG1_Chk_B_H : BOOL;  (* 【Y806】B(右側) NG1チャック戻; at IOBus://unit#8/Output Bit 32 bits/Output Bit 06 *)
    Out_CYw_NG1_Chk_B_F : BOOL;  (* 【Y807】B(右側) NG1チャック行; at IOBus://unit#8/Output Bit 32 bits/Output Bit 07 *)
    Out_CYw_Rev_01_Chk_B_H : BOOL;  (* 【Y808】B(右側)ST4 反転1チャック閉 戻; at IOBus://unit#8/Output Bit 32 bits/Output Bit 08 *)
    Out_CYw_Rev_01_Chk_B_F : BOOL;  (* 【Y809】B(右側)ST4 反転1チャック開 戻; at IOBus://unit#8/Output Bit 32 bits/Output Bit 09 *)
    Out_CYw_Rev_01_Pick_B_H : BOOL;  (* 【Y810】B(右側)ST4 反転1ピックアップ戻; at IOBus://unit#8/Output Bit 32 bits/Output Bit 10 *)
    Out_CYw_Rev_01_Pick_B_F : BOOL;  (* 【Y811】B(右側)ST4 反転1ピックアップ行; at IOBus://unit#8/Output Bit 32 bits/Output Bit 11 *)
    Out_CYw_Rev_02_Chk_B_H : BOOL;  (* 【Y812】B(右側)ST6 反転2チャック閉 戻; at IOBus://unit#8/Output Bit 32 bits/Output Bit 12 *)
    Out_CYw_Rev_02_Chk_B_F : BOOL;  (* 【Y813】B(右側)ST6 反転2チャック開 行; at IOBus://unit#8/Output Bit 32 bits/Output Bit 13 *)
    Out_CYw_Rev_02_Pick_B_H : BOOL;  (* 【Y814】B(右側)ST6 反転2ピックアップ戻; at IOBus://unit#8/Output Bit 32 bits/Output Bit 14 *)
    Out_CYw_Rev_02_Pick_B_F : BOOL;  (* 【Y815】B(右側)ST6 反転2ピックアップ行; at IOBus://unit#8/Output Bit 32 bits/Output Bit 15 *)
    Out_CYw_Disc_Chk_B_H : BOOL;  (* 【Y816】B(右側) 排出チャック閉 戻; at IOBus://unit#8/Output Bit 32 bits/Output Bit 16 *)
    Out_CYw_Disc_Chk_B_F : BOOL;  (* 【Y817】B(右側) 排出チャック開 行; at IOBus://unit#8/Output Bit 32 bits/Output Bit 17 *)
    Out_CYw_Ejc_Hldr_Feed_B_F : BOOL;  (* 【Y819】B(右側) 排出フォルダ送り行; at IOBus://unit#8/Output Bit 32 bits/Output Bit 19 *)
    Out_CYw_Ejc_Hldr_Feed_B_H : BOOL;  (* 【Y818】B(右側) 排出フォルダ送り戻; at IOBus://unit#8/Output Bit 32 bits/Output Bit 18 *)
    Out_CYS_Pos_01_Stopper_B : BOOL;  (* 【Y820】B(右側) 位置1ストッパー; at IOBus://unit#8/Output Bit 32 bits/Output Bit 20 *)
    Out_CYS_Pos_02_Stopper_B : BOOL;  (* 【Y821】B(右側) 位置2ストッパー; at IOBus://unit#8/Output Bit 32 bits/Output Bit 21 *)
    Out_CYS_Pos_03_Stopper_B : BOOL;  (* 【Y822】B(右側) 位置3ストッパー; at IOBus://unit#8/Output Bit 32 bits/Output Bit 22 *)
    Out_CYS_Pos_04_Stopper_B : BOOL;  (* 【Y823】B(右側) 位置4ストッパー; at IOBus://unit#8/Output Bit 32 bits/Output Bit 23 *)
    Out_CYS_Pos_05_Stopper_B : BOOL;  (* 【Y824】B(右側) 位置5ストッパー; at IOBus://unit#8/Output Bit 32 bits/Output Bit 24 *)
    Out_CYS_Pos_06_Stopper_B : BOOL;  (* 【Y825】B(右側) 位置6ストッパー; at IOBus://unit#8/Output Bit 32 bits/Output Bit 25 *)
    Out_CYw_SH_B_Turn_H : BOOL;  (* 【Y826】B(右側) ストックフォルダターン戻; at IOBus://unit#8/Output Bit 32 bits/Output Bit 26 *)
    Out_CYw_SH_B_Turn_F : BOOL;  (* 【Y827】B(右側) ストックフォルダターン行; at IOBus://unit#8/Output Bit 32 bits/Output Bit 27 *)
    Out_CYw_NG1_Srt_B_H : BOOL;  (* 【Y828】B(右側) NG1仕分け 戻; at IOBus://unit#8/Output Bit 32 bits/Output Bit 28 *)
    Out_CYw_NG1_Srt_B_F : BOOL;  (* 【Y829】B(右側) NG1仕分け 行; at IOBus://unit#8/Output Bit 32 bits/Output Bit 29 *)
    TimerQ_In_Sen_Accum_CV_A_Full : BOOL;  (* 【X200】A(左側) アキュームA() CV満 *)
    TimerQ_In_Sen_Accum_CV_A_Arrival : BOOL;  (* 【X201】A(左側) アキュームA ()CV着 *)
    TimerQ_In_Sen_Work_A_Pos_00 : BOOL;  (* 【X202】A(左側)ワーク位置0 *)
    TimerQ_In_Sen_Work_A_Pos_01 : BOOL;  (* 【X203】A(左側)ワーク位置1 *)
    TimerQ_In_Sen_Work_A_Pos_02 : BOOL;  (* 【X204】A(左側)ワーク位置2 *)
    TimerQ_In_Sen_Work_A_Pos_03 : BOOL;  (* 【X205】A(左側)ワーク位置3 *)
    TimerQ_In_Sen_Work_A_Pos_04 : BOOL;  (* 【X206】A(左側)ワーク位置4 *)
    TimerQ_In_Sen_Work_A_Pos_05 : BOOL;  (* 【X207】A(左側)ワーク位置5 *)
    TimerQ_In_Sen_Work_A_Pos_06 : BOOL;  (* 【X208】A(左側)ワーク位置6 *)
    TimerQ_In_Sen_Work_A_Pos_07 : BOOL;  (* 【X209】A(左側)ワーク位置7 *)
    TimerQ_In_Sen_NG1_Tray_01_A_Full : BOOL;  (* 【X210】A(左側) NG1トレイ1満杯 *)
    TimerQ_In_Sen_NG1_Tray_01_A_Full_Warn : BOOL;  (* 【X211】A(左側) NG1トレイ1満杯警告 *)
    TimerQ_In_Sen_NG1_Tray_02_A_Full : BOOL;  (* 【X212】A(左側) NG1トレイ2満杯停止 *)
    TimerQ_In_Sen_NG1_Tray_02_A_Full_Warn : BOOL;  (* 【X213】A(左側) NG1トレイ2満杯警告 *)
    TimerQ_In_Sen_SH_A_Ent : BOOL;  (* 【X214】A(左側) ストックフォルダIN *)
    TimerQ_In_Sen_SH_A_Ext : BOOL;  (* 【X215】A(左側) ストックフォルダOut *)
    TimerQ_In_Sen_SH_A_Type_Ent : BOOL;  (* 【X216】A(左側) ストック機種判別IN *)
    TimerQ_In_Sen_SH_A_Type_Ext : BOOL;  (* 【X217】A(左側) ストック機種判別OUT *)
    TimerQ_In_SenCY_Sply_Slide_A_H : BOOL;  (* 【X218】A(左側) 供給スライド戻 *)
    TimerQ_In_SenCY_Sply_Slide_A_F : BOOL;  (* 【X219】A(左側) 供給スライド行 *)
    TimerQ_In_SenCY_Sply_Pick_A_H : BOOL;  (* 【X220】A(左側) 供給ピックアップ戻 *)
    TimerQ_In_SenCY_Sply_Pick_A_F : BOOL;  (* 【X221】A(左側) 供給ピックアップ行 *)
    TimerQ_In_SenCY_Sply_Chk_A_H : BOOL;  (* 【X222】A(左側) 供給チャック戻 *)
    TimerQ_In_SenCY_Sply_Chk_A_F : BOOL;  (* 【X223】A(左側) 供給チャック行 *)
    TimerQ_In_SenCY_HgtInsp_Clp_A_H : BOOL;  (* 【X224】A(左側) 高さ検査押え戻 *)
    TimerQ_In_SenCY_HgtInsp_Clp_A_F : BOOL;  (* 【X225】A(左側) 高さ検査押え行 *)
    TimerQ_In_SenCY_HgtInsp_Lf_A_H : BOOL;  (* 【X226】A(左側) 高さ検査持上戻 *)
    TimerQ_In_SenCY_HgtInsp_Lf_A_F : BOOL;  (* 【X227】A(左側) 高さ検査持上行 *)
    TimerQ_In_SenCY_NG1_Pick_A_H : BOOL;  (* 【X228】A(左側) NG1ピックアップ戻 *)
    TimerQ_In_SenCY_NG1_Pick_A_F : BOOL;  (* 【X229】A(左側) NG1ピックアップ行 *)
    TimerQ_In_SenCY_NG1_Chk_A_H : BOOL;  (* 【X230】A(左側) NG1チャック戻 *)
    TimerQ_In_SenCY_NG1_Chk_A_F : BOOL;  (* 【X231】A(左側) NG1チャック行 *)
    TimerQ_In_SenCY_Rev_01_Chk_A_H : BOOL;  (* 【X300】A(左側)ST4 反転1チャック戻 *)
    TimerQ_In_SenCY_Rev_01_Chk_A_F : BOOL;  (* 【X301】A(左側)ST4 反転1チャック行 *)
    TimerQ_In_SenCY_Rev_01_Pick_A_H : BOOL;  (* 【X302】A(左側)ST4 反転1ピックアップ戻 *)
    TimerQ_In_SenCY_Rev_01_Pick_A_F : BOOL;  (* 【X303】A(左側)ST4 反転1ピックアップ行 *)
    TimerQ_In_SenCY_Rev_02_Chk_A_H : BOOL;  (* 【X304】A(左側)ST6 反転2チャック戻 *)
    TimerQ_In_SenCY_Rev_02_Chk_A_F : BOOL;  (* 【X305】A(左側)ST6 反転2チャック行 *)
    TimerQ_In_SenCY_Rev_02_Pick_A_H : BOOL;  (* 【X306】A(左側)ST6 反転2ピックアップ戻 *)
    TimerQ_In_SenCY_Rev_02_Pick_A_F : BOOL;  (* 【X307】A(左側)ST6 反転2ピックアップ行 *)
    TimerQ_In_SenCY_Disc_Chk_A_H : BOOL;  (* 【X308】A(左側) 排出チャック戻 *)
    TimerQ_In_SenCY_Disc_Chk_A_F : BOOL;  (* 【X309】A(左側) 排出チャック行 *)
    TimerQ_In_SenCY_Ejc_SH_Feed_A_H : BOOL;  (* 【X310】A(左側) 排出フォルダ送り戻 *)
    TimerQ_In_SenCY_Ejc_SH_Feed_A_F : BOOL;  (* 【X311】A(左側) 排出フォルダ送り行 *)
    TimerQ_In_SenCY_Pos_01_Stopper_A_H : BOOL;  (* 【X312】A(左側) 位置1ストッパー戻 *)
    TimerQ_In_SenCY_Pos_01_Stopper_A_F : BOOL;  (* 【X313】位置1ストッパー行 *)
    TimerQ_In_SenCY_Pos_02_Stopper_A_H : BOOL;  (* 【X314】A(左側) 位置2ストッパー戻 *)
    TimerQ_In_SenCY_Pos_02_Stopper_A_F : BOOL;  (* 【X315】A(左側) 位置2ストッパー行 *)
    TimerQ_In_SenCY_Pos_03_Stopper_A_H : BOOL;  (* 【X316】A(左側) 位置3ストッパー戻 *)
    TimerQ_In_SenCY_Pos_03_Stopper_A_F : BOOL;  (* 【X317】A(左側) 位置3ストッパー行 *)
    TimerQ_In_SenCY_Pos_04_Stopper_A_H : BOOL;  (* 【X318】A(左側) 位置4ストッパー戻 *)
    TimerQ_In_SenCY_Pos_04_Stopper_A_F : BOOL;  (* 【X319】A(左側) 位置4ストッパー行 *)
    TimerQ_In_SenCY_Pos_05_Stopper_A_H : BOOL;  (* 【X320】A(左側) 位置5ストッパー戻 *)
    TimerQ_In_SenCY_Pos_05_Stopper_A_F : BOOL;  (* 【X321】A(左側) 位置5ストッパー行 *)
    TimerQ_In_SenCY_Pos_06_Stopper_A_H : BOOL;  (* 【X322】A(左側) 位置6ストッパー戻 *)
    TimerQ_In_SenCY_Pos_06_Stopper_A_F : BOOL;  (* 【X323】A(左側) 位置6ストッパー行 *)
    TimerQ_In_SenCY_SH_A_Turn_H : BOOL;  (* 【X324】A(左側) ストックフォルダターン戻 *)
    TimerQ_In_SenCY_SH_A_Turn_F : BOOL;  (* 【X325】A(左側) ストックフォルダターン行 *)
    TimerQ_In_SenCY_NG1_Srt_A_H : BOOL;  (* 【X330】NG1仕分け 戻 *)
    TimerQ_In_SenCY_NG1_Srt_A_F : BOOL;  (* 【X331】NG1仕分け 行 *)
    TimerQ_In_Sen_Accum_CV_B_Full : BOOL;  (* 【X400】B(右側) アキュームCV満 *)
    TimerQ_In_Sen_Accum_CV_B_Arrival : BOOL;  (* 【X401】B(右側) アキュームCV着 *)
    TimerQ_In_Sen_Work_B_Pos_00 : BOOL;  (* 【X402】B(右側)ワーク位置0 *)
    TimerQ_In_Sen_Work_B_Pos_01 : BOOL;  (* 【X403】B(右側)ワーク位置1 *)
    TimerQ_In_Sen_Work_B_Pos_02 : BOOL;  (* 【X404】B(右側)ワーク位置2 *)
    TimerQ_In_Sen_Work_B_Pos_03 : BOOL;  (* 【X405】B(右側)ワーク位置3 *)
    TimerQ_In_Sen_Work_B_Pos_04 : BOOL;  (* 【X406】B(右側)ワーク位置4 *)
    TimerQ_In_Sen_Work_B_Pos_05 : BOOL;  (* 【X407】B(右側)ワーク位置5 *)
    TimerQ_In_Sen_Work_B_Pos_06 : BOOL;  (* 【X408】B(右側)ワーク位置6 *)
    TimerQ_In_Sen_Work_B_Pos_07 : BOOL;  (* 【X409】B(右側)ワーク位置7 *)
    TimerQ_In_Sen_NG1_Tray_01_B_Full : BOOL;  (* 【X410】B(右側) NG1トレイ1満杯 *)
    TimerQ_In_Sen_NG1_Tray_01_B_Full_Warn : BOOL;  (* 【X411】B(右側) NG1トレイ1満杯警告 *)
    TimerQ_In_Sen_NG1_Tray_02_B_Full : BOOL;  (* 【X412】B(右側) NG1トレイ2満杯停止 *)
    TimerQ_In_Sen_NG1_Tray_02_B_Full_Warn : BOOL;  (* 【X413】B(右側) NG1トレイ2満杯警告 *)
    TimerQ_In_Sen_SH_B_Ent : BOOL;  (* 【X414】B(右側) ストックフォルダIN *)
    TimerQ_In_Sen_SH_B_Ext : BOOL;  (* 【X415】B(右側) ストックフォルダOut *)
    TimerQ_In_Sen_SH_B_Type_Ent : BOOL;  (* 【X416】B(右側) ストック機種判別IN *)
    TimerQ_In_Sen_SH_B_Type_Ext : BOOL;  (* 【X417】B(右側) ストック機種判別OUT *)
    TimerQ_In_SenCY_Sply_Slide_B_H : BOOL;  (* 【X418】B(右側) 供給スライド戻 *)
    TimerQ_In_SenCY_Sply_Slide_B_F : BOOL;  (* 【X419】B(右側) 供給スライド行 *)
    TimerQ_In_SenCY_Sply_Pick_B_H : BOOL;  (* 【X420】B(右側) 供給ピックアップ戻 *)
    TimerQ_In_SenCY_Sply_Pick_B_F : BOOL;  (* 【X421】B(右側) 供給ピックアップ行 *)
    TimerQ_In_SenCY_Sply_Chk_B_H : BOOL;  (* 【X422】B(右側) 供給チャック閉 戻 *)
    TimerQ_In_SenCY_HgtInsp_Clp_B_H : BOOL;  (* 【X424】B(右側) 高さ検査押え戻 *)
    TimerQ_In_SenCY_Sply_Chk_B_F : BOOL;  (* 【X423】B(右側) 供給チャック開 行 *)
    TimerQ_In_SenCY_HgtInsp_Clp_B_F : BOOL;  (* 【X425】B(右側) 高さ検査押え行 *)
    TimerQ_In_SenCY_HgtInsp_Lf_B_H : BOOL;  (* 【X426】B(右側) 高さ検査持上戻 *)
    TimerQ_In_SenCY_HgtInsp_Lf_B_F : BOOL;  (* 【X427】 B(右側) 高さ検査持上行 *)
    TimerQ_In_SenCY_NG1_Pick_B_H : BOOL;  (* 【X428】B(右側) NG1ピックアップ戻 *)
    TimerQ_In_SenCY_NG1_Pick_B_F : BOOL;  (* 【X429】B(右側) NG1ピックアップ行 *)
    TimerQ_In_SenCY_NG1_Chk_B_H : BOOL;  (* 【X430】 B(右側) NG1チャック閉 戻 *)
    TimerQ_In_SenCY_NG1_Chk_B_F : BOOL;  (* 【X431】B(右側) NG1チャック開 行 *)
    TimerQ_In_SenCY_Rev_01_Chk_B_H : BOOL;  (* 【X500】B(右側)ST4 反転1チャック閉 戻 *)
    TimerQ_In_SenCY_Rev_01_Pick_B_H : BOOL;  (* 【X502】B(右側)ST4 反転1ピックアップ戻 *)
    TimerQ_In_SenCY_Rev_01_Pick_B_F : BOOL;  (* 【X503】B(右側)ST4 反転1ピックアップ行 *)
    TimerQ_In_SenCY_Rev_02_Chk_B_H : BOOL;  (* 【X504】B(右側)ST6 反転2チャック閉 戻 *)
    TimerQ_In_SenCY_Rev_02_Chk_B_F : BOOL;  (* 【X505】B(右側)ST6 反転2チャック開 行 *)
    TimerQ_In_SenCY_Rev_02_Pick_B_H : BOOL;  (* 【X506】B(右側)ST6 反転2ピックアップ戻 *)
    TimerQ_In_SenCY_Rev_02_Pick_B_F : BOOL;  (* 【X507】B(右側)ST6 反転2ピックアップ行 *)
    TimerQ_In_SenCY_Disc_Chk_B_H : BOOL;  (* 【X508】B(右側) 排出チャック閉 戻 *)
    TimerQ_In_SenCY_Disc_Chk_B_F : BOOL;  (* 【X509】B(右側) 排出チャック開 行 *)
    TimerQ_In_SenCY_Ejc_SH_Feed_B_H : BOOL;  (* 【X511】B(右側) 排出フォルダ送り行 *)
    TimerQ_In_SenCY_Ejc_SH_Feed_B_F : BOOL;  (* 【X510】B(右側) 排出フォルダ送り戻 *)
    TimerQ_In_SenCY_Pos_01_Stopper_B_H : BOOL;  (* 【X512】B(右側) 位置1ストッパー戻 *)
    TimerQ_In_SenCY_Pos_01_Stopper_B_F : BOOL;  (* 【X513】B(右側) 位置1ストッパー行 *)
    TimerQ_In_SenCY_Pos_02_Stopper_B_H : BOOL;  (* 【X514】B(右側) 位置2ストッパー戻 *)
    TimerQ_In_SenCY_Pos_02_Stopper_B_F : BOOL;  (* 【X515】B(右側) 位置2ストッパー行 *)
    TimerQ_In_SenCY_Pos_03_Stopper_B_H : BOOL;  (* 【X516】B(右側) 位置3ストッパー戻 *)
    TimerQ_In_SenCY_Pos_03_Stopper_B_F : BOOL;  (* 【X517】B(右側) 位置3ストッパー行 *)
    TimerQ_In_SenCY_Pos_04_Stopper_B_H : BOOL;  (* 【X518】B(右側) 位置4ストッパー戻 *)
    TimerQ_In_SenCY_Pos_04_Stopper_B_F : BOOL;  (* 【X519】B(右側) 位置4ストッパー行 *)
    TimerQ_In_SenCY_Pos_05_Stopper_B_H : BOOL;  (* 【X520】B(右側) 位置5ストッパー戻 *)
    TimerQ_In_SenCY_Pos_05_Stopper_B_F : BOOL;  (* 【X521】B(右側) 位置5ストッパー行 *)
    TimerQ_In_SenCY_Pos_06_Stopper_B_H : BOOL;  (* 【X522】B(右側) 位置6ストッパー戻 *)
    TimerQ_In_SenCY_Pos_06_Stopper_B_F : BOOL;  (* 【X523】B(右側) 位置6ストッパー行 *)
    TimerQ_In_SenCY_SH_B_Turn_H : BOOL;  (* 【X524】B(右側) ストックフォルダターン戻 *)
    TimerQ_In_SenCY_SH_B_Turn_F : BOOL;  (* 【X525】B(右側) ストックフォルダターン行 *)
    TimerQ_In_SenCY_NG1_Srt_B_H : BOOL;  (* 【X530】B(右側) NG1仕分け 戻 *)
    TimerQ_In_SenCY_NG1_Srt_B_F : BOOL;  (* 【X531】B(右側) NG1仕分け 行 *)
    TimerQ_In_Sen_Supply_Container_Exist : BOOL;  (* 【X1000】供給部コンテナ有 *)
    TimerQ_In_Sen_Destacker_Stage_01_Exist : BOOL;  (* 【X1001】段バラシ1段目有 *)
    TimerQ_In_Sen_Destacker_Stage_02_Exist : BOOL;  (* 【X1002】段バラシ2段目有 *)
    TimerQ_In_Sen_Container_Arrival : BOOL;  (* 【X1003】コンテナ到着 *)
    TimerQ_In_Sen_Container_Direction_Check : BOOL;  (* 【X1004】コンテナ方向確認 *)
    TimerQ_In_Sen_Container_Pass : BOOL;  (* 【X1005】コンテナ通過 *)
    TimerQ_In_Sen_Container_Full : BOOL;  (* 【X1006】コンテナ満杯 *)
    TimerQ_In_Sen_Container_Sorting : BOOL;  (* 【X1007】コンテナ仕分け *)
    TimerQ_In_SenCY_Empty_Container_CY_H : BOOL;  (* 【X1010】空コンテナ送り 戻 *)
    TimerQ_In_SenCY_Empty_Container_CY_F : BOOL;  (* 【X1011】空コンテナ送り 行 *)
    TimerQ_In_SenCY_Sep_Claw1_H : BOOL;  (* 【X1012】段バラシ爪1 戻 *)
    TimerQ_In_SenCY_Sep_Claw1_F : BOOL;  (* 【X1013】段バラシ爪1 行 *)
    TimerQ_In_SenCY_Sep_Claw2_F : BOOL;  (* 【X1015】段バラシ爪2 行 *)
    TimerQ_In_SenCY_Sep_Claw2_H : BOOL;  (* 【X1014】段バラシ爪2 戻 *)
    TimerQ_In_SenCY_Ejc_Cont1_H : BOOL;  (* 【X1016】コンテナ排出1 戻 *)
    TimerQ_In_SenCY_Ejc_Cont1_F : BOOL;  (* 【X1017】コンテナ排出1 行 *)
    TimerQ_In_SenCY_Ejc_Cont2_H : BOOL;  (* 【X1018】コンテナ排出2 戻 *)
    TimerQ_In_SenCY_Ejc_Cont2_F : BOOL;  (* 【X1019】コンテナ排出2 行 *)
    TimerQ_In_SenCY_Box_Chk_H : BOOL;  (* 【X1020】箱入れチャック 戻 *)
    TimerQ_In_SenCY_Box_Chk_F : BOOL;  (* 【X1021】箱入れチャック 行 *)
    TimerQ_In_SenCY_Srt_Stopper_H : BOOL;  (* 【X1022】コンテナ仕分けストッパー 戻 *)
    TimerQ_In_SenCY_Srt_Stopper_F : BOOL;  (* 【X1023】コンテナ仕分けストッパー 行 *)
    TimerQ_In_SenCY_Srt_Feed_H : BOOL;  (* 【X1024】コンテナ仕分け送り 戻 *)
    TimerQ_In_SenCY_Srt_Feed_F : BOOL;  (* 【X1025】コンテナ仕分け送り 行 *)
    TimerQ_In_Sen_Unl_Conv_A_Pass : BOOL;  (* 【X1100】A(左側) 取出しコンベア 通過 *)
    TimerQ_In_Sen_Unl_Conv_B_Pass : BOOL;  (* 【X1101】B(右側) 取出しコンベア 通過 *)
    TimerQ_In_Sen_Trs_Conv_B_Arrival : BOOL;  (* 【X1103】B(右側) 搬送コンベア到着 *)
    TimerQ_In_Sen_Trs_Conv_A_Arrival : BOOL;  (* 【X1102】A(左側) 搬送コンベア到着 *)
    TimerQ_In_SenCY_Hnd_Feed_A_H : BOOL;  (* 【X1104】A(左側) コンベア受渡送り戻 *)
    TimerQ_In_SenCY_Hnd_Feed_A_F : BOOL;  (* 【X1105】A(左側) コンベア受渡送り行 *)
    TimerQ_In_SenCY_Hnd_Feed_B_H : BOOL;  (* 【X1106】B(右側) コンベア受渡送り戻 *)
    TimerQ_In_SenCY_Hnd_Feed_B_F : BOOL;  (* 【X1107】B(右側) コンベア受渡送り行 *)
    TimerQ_In_SenCY_Rev_01_Chk_B_F : BOOL;  (* 【X501】B(右側)ST4 反転1チャック開 行 *)
    AutoMode : BOOL;  (* 自動運転 *)
    ManualMode : BOOL;  (* 手動運転 *)
    M9999 : BOOL;  (* 非常停止 *)
    Out_CYw_Sply_Slide_A_H_Done : BOOL;  (* 【Y616】A(左側) 供給スライド戻 動作完了 *)
END_VAR
VAR_GLOBAL RETAIN
    Output_A_Error_M : ARRAY[0..99] OF Bool;  (* A(左側)出力 エラー：; [1] 【Y616】A(左側) 供給スライド戻; [2] 【Y617】A(左側) 供給スライド行; [3] 【Y618】A(左側) 供給ピックアップ戻; [4] 【Y619】A(左側) 供給ピックアップ行; [5] 【Y620】A(左側) 供給チャック閉 戻; [6] 【Y621】A(左側) 供給チャック開 行; [7] 【Y700】A(左側) 高さ検査押え戻; [8] 【Y701】A(左側) 高さ検査押え行; [9] 【Y702】A(左側) 高さ検査持上戻; [10] 【Y703】A(左側) 高さ検査持上行; [11] 【Y704】A(左側) NG1ピックアップ戻; [12] 【Y705】A(左側) NG1ピックアップ 行; [13] 【Y706】A(左側) NG1チャック戻; [14] 【Y707】A(左側) NG1チャック行; [15] 【Y708】A(左側)ST4 反転1チャック閉; [16] 【Y709】A(左側)ST4 反転1チャック開; [17] 【Y710】A(左側)ST4 反転1ピックアップ戻; [18] 【Y711】A(左側)ST4 反転1ピックアップ行; [19] 【Y712】A(左側)ST6 反転2チャック閉 戻; [20] 【Y713】A(左側)ST6 反転2チャック開 行; [21] 【Y714】A(左側)ST6 反転2ピックアップ戻; [22] 【Y715】A(左側)ST6 反転2ピックアップ行; [23] 【Y716】A(左側) 排出チャック閉 戻; [24] 【Y717】A(左側) 排出チャック開 行; [25] 【Y718】A(左側) 排出フォルダ送り戻; [26] 【Y719】A(左側) 排出フォルダ送り行; [27] A(左側) 位置1ストッパー戻; [28] 【Y720】A(左側) 位置1ストッパー 行; [29] 【Y721】A(左側) 位置2ストッパー; [30] 【Y721】A(左側) 位置2ストッパー; [31] 【Y722】A(左側) 位置3ストッパー戻; [32] 【Y722】A(左側) 位置3ストッパー行; [34] 【Y723】A(左側) 位置4ストッパー行; [35] 【Y724】A(左側) 位置5ストッパー戻; [36] 【Y724】A(左側) 位置5ストッパー行; [37] 【Y725】A(左側) 位置6ストッパー戻; [38] 【Y725】A(左側) 位置6ストッパー行; [39] 【Y726】A(左側) ストックフォルダターン戻; [40] 【Y727】A(左側) ストックフォルダターン行; [41] 【Y728】A(左側) NG1仕分け 戻; [42] 【Y729】A(左側) NG1仕分け 行; [43] 【Y1300】A(左側) コンベア受渡送り戻; [44] 【Y1301】A(左側) コンベア受渡送り行 *)
    Output_A_Restart_M : ARRAY[0..99] OF Bool;  (* A(左側)出力 再スタート：; [1] 【Y616】A(左側) 供給スライド戻; [2] 【Y617】A(左側) 供給スライド行; [3] 【Y618】A(左側) 供給ピックアップ戻; [4] 【Y619】A(左側) 供給ピックアップ行; [5] 【Y620】A(左側) 供給チャック閉 戻; [6] 【Y621】A(左側) 供給チャック開 行; [7] 【Y700】A(左側) 高さ検査押え戻; [8] 【Y701】A(左側) 高さ検査押え行; [9] 【Y702】A(左側) 高さ検査持上戻; [10] 【Y703】A(左側) 高さ検査持上行; [11] 【Y704】A(左側) NG1ピックアップ戻; [12] 【Y705】A(左側) NG1ピックアップ 行; [13] 【Y706】A(左側) NG1チャック戻; [14] 【Y707】A(左側) NG1チャック行; [15] 【Y708】A(左側)ST4 反転1チャック閉; [16] 【Y709】A(左側)ST4 反転1チャック開; [17] 【Y710】A(左側)ST4 反転1ピックアップ戻; [18] 【Y711】A(左側)ST4 反転1ピックアップ行; [19] 【Y712】A(左側)ST6 反転2チャック閉 戻; [20] 【Y713】A(左側)ST6 反転2チャック開 行; [21] 【Y714】A(左側)ST6 反転2ピックアップ戻; [22] 【Y715】A(左側)ST6 反転2ピックアップ行; [23] 【Y716】A(左側) 排出チャック閉 戻; [24] 【Y717】A(左側) 排出チャック開 行; [25] 【Y718】A(左側) 排出フォルダ送り戻; [26] 【Y719】A(左側) 排出フォルダ送り行; [27] A(左側) 位置1ストッパー戻; [28] 【Y720】A(左側) 位置1ストッパー 行; [29] 【Y721】A(左側) 位置2ストッパー; [30] 【Y721】A(左側) 位置2ストッパー; [31] 【Y722】A(左側) 位置3ストッパー戻; [32] 【Y722】A(左側) 位置3ストッパー行; [34] 【Y723】A(左側) 位置4ストッパー行; [35] 【Y724】A(左側) 位置5ストッパー戻; [36] 【Y724】A(左側) 位置5ストッパー行; [37] 【Y725】A(左側) 位置6ストッパー戻; [38] 【Y725】A(左側) 位置6ストッパー行; [39] 【Y726】A(左側) ストックフォルダターン戻; [40] 【Y727】A(左側) ストックフォルダターン行; [41] 【Y728】A(左側) NG1仕分け 戻; [42] 【Y729】A(左側) NG1仕分け 行; [43] 【Y1300】A(左側) コンベア受渡送り戻; [44] 【Y1301】A(左側) コンベア受渡送り行 *)
END_VAR
VAR_GLOBAL
    Out_SW_Start_LP_GREEN_Auto : ARRAY[0..10] OF Bool;  (* 自動 【Y600】SWスタートランプ緑：; [1] 1 *)
    Out_SW_Start_LP_GREEN_Manual : ARRAY[0..10] OF Bool;  (* 手動 【Y600】SWスタートランプ緑： *)
    Out_SW_Stop_LP_RED_Auto : ARRAY[0..10] OF Bool;  (* 【Y601】SWストップランプ赤： *)
    Out_SW_Stop_LP_RED_Manual : ARRAY[0..10] OF Bool;  (* 【Y601】SWストップランプ赤： *)
    Out_SW_Reset_LP_Orange_Auto : ARRAY[0..10] OF Bool;  (* 【Y602】SW リセットランプ橙： *)
    Out_SW_Reset_LP_Orange_Manual : ARRAY[0..10] OF Bool;  (* 【Y602】SW リセットランプ橙： *)
    Out_Sg_LP_GREEN_Auto : ARRAY[0..10] OF Bool;  (* 【Y603】シグナルタワー緑： *)
    Out_Sg_LP_GREEN_Manual : ARRAY[0..10] OF Bool;  (* 【Y603】シグナルタワー緑： *)
    Out_Sg_LP_RED_Auto : ARRAY[0..10] OF Bool;  (* 【Y604】シグナルタワー赤： *)
    Out_Sg_LP_RED_Manual : ARRAY[0..10] OF Bool;  (* 【Y604】シグナルタワー赤： *)
    Out_Sg_LP_ORANGE_Auto : ARRAY[0..10] OF Bool;  (* 【Y605】シグナルタワー橙： *)
    Out_Sg_LP_ORANGE_Manual : ARRAY[0..10] OF Bool;  (* 【Y605】シグナルタワー橙： *)
    Out_Sg_BUZZER_Auto : ARRAY[0..10] OF Bool;  (* 【Y606】シグナルタワーブザー： *)
    Out_Sg_BUZZER_Manual : ARRAY[0..10] OF Bool;  (* 【Y606】シグナルタワーブザー： *)
    Out_Accum_Cv_RESET_Manual : ARRAY[0..10] OF Bool;  (* 【Y608】アキューム コンベア リセット： *)
    Out_Accum_Cv_RESET_Auto : ARRAY[0..10] OF Bool;  (* 【Y608】アキューム コンベア リセット： *)
    Out_Acc_Conv_Run_Manual : ARRAY[0..10] OF Bool;  (* 【Y607】アキューム コンベア運転ON： *)
    Out_Acc_Conv_Run_Auto : ARRAY[0..10] OF Bool;  (* 【Y607】アキューム コンベア運転ON： *)
    Out_Accum_Cv_PowerOn_Auto : ARRAY[0..10] OF Bool;  (* 【Y609】アキューム コンベア電源ON： *)
    Out_Accum_Cv_PowerOn_Manual : ARRAY[0..10] OF Bool;  (* 【Y609】アキューム コンベア電源ON： *)
    Out_Insp_Cv_A_Run_Auto : ARRAY[0..10] OF Bool;  (* 【Y610】A(左側) 検査 コンベア運転ON： *)
    Out_Insp_Cv_A_Run_Manual : ARRAY[0..10] OF Bool;  (* 【Y610】A(左側) 検査 コンベア運転ON： *)
    Out_Insp_Cv_A_RESET_Auto : ARRAY[0..10] OF Bool;  (* 【Y611】A(左側) 検査 コンベア リセット： *)
    Out_Insp_Cv_A_RESET_Manual : ARRAY[0..10] OF Bool;  (* 【Y611】A(左側) 検査 コンベア リセット： *)
    Out_Insp_Cv_A_PowerOn_Auto : ARRAY[0..10] OF Bool;
    Out_Insp_Cv_A_PowerOn_Manual : ARRAY[0..10] OF Bool;
    Out_Insp_Cv_B_RESET_Auto : ARRAY[0..10] OF Bool;  (* 【Y614】B(右側) 検査 コンベア リセット： *)
    Out_Insp_Cv_B_RESET_Manual : ARRAY[0..10] OF Bool;  (* 【Y614】B(右側) 検査 コンベア リセット： *)
    Out_Insp_Cv_B_Run_Manual : ARRAY[0..10] OF Bool;  (* 【Y613】B(右側) 検査 コンベア運転ON： *)
    Out_Insp_Cv_B_Run_Auto : ARRAY[0..10] OF Bool;  (* 【Y613】B(右側) 検査 コンベア運転ON： *)
    Out_CYw_Sply_Slide_A_H_Manual : ARRAY[0..10] OF Bool;  (* 手動【Y616】A(左側) 供給スライド戻： *)
    Out_CYw_Sply_Slide_A_H_Auto : ARRAY[0..10] OF Bool;  (* 自動【Y616】A(左側) 供給スライド戻：; [1] 原点位置移動; [2] ワーク設置完了後 *)
    HMI_MessageNo : ARRAY[0..9] OF UINT;  (* メッセージNo *)
    HMI_Message : ARRAY[0..9] OF String[256];  (* メッセージ内容 *)
    HMI_Language : BOOL;  (* 言語切替 *)
    Out_CYw_Sply_Slide_A_F_Done : BOOL;  (* 【Y617】A(左側) 供給スライド行動作完了 *)
    Pause : ARRAY[0..99] OF Bool;  (* 一時停止：; [1] シリンダ; [2] コンベア＆ドアセンサ; [3] FH A(左側) ST1; [4] A(左側)検査コンベア ワーク不一致; [5] PCON1 1; [6] GT2 エラー; [7] NG1仕分けエラー; [8] 反転1エラー; [9] FH A(左側) ST5; [10] FH B(右側) ST1; [11] FH B(右側) ST5; [12] A(左側) ST6 反転2 ワーク不一致 *)
END_VAR
VAR_GLOBAL RETAIN
    Output_B_Error_M : ARRAY[0..99] OF Bool;  (* B(右側)出力 エラー：; [1] 【Y622】B(右側) 供給スライド戻; [2] 【Y623】B(右側) 供給スライド行; [3] 【Y624】B(右側) 供給ピックアップ戻; [4] 【Y625】B(右側) 供給ピックアップ行; [5] 【Y626】B(右側) 供給チャック閉 戻; [6] 【Y627】B(右側) 供給チャック開 行; [7] 【Y800】B(右側) 高さ検査押え戻; [9] 【Y802】B(右側) 高さ検査持上戻; [11] 【Y804】B(右側) NG1ピックアップ戻; [12] 【Y805】B(右側) NG1ピックアップ 行; [14] 【Y807】B(右側) NG1チャック行; [18] 【Y811】B(右側)ST4 反転1ピックアップ行; [23] 【Y816】B(右側) 排出チャック閉 戻; [42] 【Y829】B(右側) NG1仕分け 行; [41] 【Y828】B(右側) NG1仕分け 戻; [40] 【Y827】B(右側) ストックフォルダターン行; [39] 【Y826】B(右側) ストックフォルダターン戻; [38] 【Y825】B(右側) 位置6ストッパー行; [37] 【Y825】B(右側) 位置6ストッパー戻; [36] 【Y824】B(右側) 位置5ストッパー行; [35] 【Y824】B(右側) 位置5ストッパー戻; [34] 【Y823】B(右側) 位置4ストッパー行; [33] 【Y823】B(右側) 位置4ストッパー戻; [32] 【Y822】B(右側) 位置3ストッパー行; [31] 【Y822】B(右側) 位置3ストッパー戻; [30] 【Y821】B(右側) 位置2ストッパー行; [29] 【Y821】B(右側) 位置2ストッパー戻; [28] 【Y820】B(右側) 位置1ストッパー 行; [27] 【Y820】B(右側) 位置1ストッパー 戻; [26] 【Y819】B(右側) 排出フォルダ送り行; [25] 【Y818】B(右側) 排出フォルダ送り戻; [24] 【Y817】B(右側) 排出チャック開 行; [22] 【Y815】B(右側)ST6 反転2ピックアップ行; [21] 【Y814】B(右側)ST6 反転2ピックアップ戻; [20] 【Y813】B(右側)ST6 反転2チャック開 行; [19] 【Y812】B(右側)ST6 反転2チャック閉 戻; [17] 【Y810】B(右側)ST4 反転1ピックアップ戻; [16] 【Y809】B(右側)ST4 反転1チャック開 戻; [15] 【Y808】B(右側)ST4 反転1チャック閉 戻; [13] 【Y806】B(右側) NG1チャック戻; [10] 【Y803】B(右側) 高さ検査持上行; [8] 【Y801】B(右側) 高さ検査押え行; [43] 【Y1302】B(右側) コンベア受渡送り戻; [44] 【Y1303】B(右側) コンベア受渡送り行 *)
    Output_B_Restart_M : ARRAY[0..99] OF Bool;  (* B(右側)出力 再スタート：; [2] 【Y623】B(右側) 供給スライド行; [3] 【Y624】B(右側) 供給ピックアップ戻; [4] 【Y625】B(右側) 供給ピックアップ行; [5] 【Y626】B(右側) 供給チャック閉 戻; [6] 【Y627】B(右側) 供給チャック開 行; [7] 【Y800】B(右側) 高さ検査押え戻; [9] 【Y802】B(右側) 高さ検査持上戻; [11] 【Y804】B(右側) NG1ピックアップ戻; [12] 【Y805】B(右側) NG1ピックアップ 行; [14] 【Y807】B(右側) NG1チャック行; [18] 【Y811】B(右側)ST4 反転1ピックアップ行; [42] 【Y829】B(右側) NG1仕分け 行; [41] 【Y828】B(右側) NG1仕分け 戻; [40] 【Y827】B(右側) ストックフォルダターン行; [39] 【Y826】B(右側) ストックフォルダターン戻; [38] 【Y825】B(右側) 位置6ストッパー行; [37] 【Y825】B(右側) 位置6ストッパー戻; [36] 【Y824】B(右側) 位置5ストッパー行; [35] 【Y824】B(右側) 位置5ストッパー戻; [34] 【Y823】B(右側) 位置4ストッパー行; [33] 【Y823】B(右側) 位置4ストッパー戻; [32] 【Y822】B(右側) 位置3ストッパー行; [31] 【Y822】B(右側) 位置3ストッパー戻; [30] 【Y821】B(右側) 位置2ストッパー行; [29] 【Y821】B(右側) 位置2ストッパー戻; [28] 【Y820】B(右側) 位置1ストッパー 行; [27] 【Y820】B(右側) 位置1ストッパー 戻; [26] 【Y819】B(右側) 排出フォルダ送り行; [25] 【Y818】B(右側) 排出フォルダ送り戻; [24] 【Y817】B(右側) 排出チャック開 行; [23] 【Y816】B(右側) 排出チャック閉 戻; [22] 【Y815】B(右側)ST6 反転2ピックアップ行; [21] 【Y814】B(右側)ST6 反転2ピックアップ戻; [20] 【Y813】B(右側)ST6 反転2チャック開 行; [19] 【Y812】B(右側)ST6 反転2チャック閉 戻; [17] 【Y810】B(右側)ST4 反転1ピックアップ戻; [16] 【Y809】B(右側)ST4 反転1チャック開 戻; [15] 【Y808】B(右側)ST4 反転1チャック閉 戻; [13] 【Y806】B(右側) NG1チャック戻; [10] 【Y803】B(右側) 高さ検査持上行; [8] 【Y801】B(右側) 高さ検査押え行; [43] 【Y1302】B(右側) コンベア受渡送り戻; [44] 【Y1303】B(右側) コンベア受渡送り行 *)
    Output_Share_Restart_M : ARRAY[0..99] OF Bool;  (* 共有出力 エラー：; [1] 【Y1200】空コンテナ送り 戻; [2] 【Y1201】空コンテナ送り 行; [3] 【Y1202】段バラシ爪 戻; [4] 【Y1203】段バラシ爪 行; [5] 【Y1204】コンテナ排出 戻; [6] 【Y1205】コンテナ排出 行; [7] 【Y1206】箱入れチャック 戻; [8] 【Y1207】箱入れチャック 行; [9] 【Y1208】コンテナ仕分けストッパー 戻; [10] 【Y1209】コンテナ仕分けストッパー 行; [11] 【Y1210】コンテナ仕分け送り 戻 *)
    Output_Share_Error_M : ARRAY[0..99] OF Bool;  (* 共有出力 再スタート：; [1] 【Y1200】空コンテナ送り 戻; [2] 【Y1201】空コンテナ送り 行; [3] 【Y1202】段バラシ爪 戻; [4] 【Y1203】段バラシ爪 行; [5] 【Y1204】コンテナ排出 戻; [6] 【Y1205】コンテナ排出 行; [8] 【Y1207】箱入れチャック 行; [9] 【Y1208】コンテナ仕分けストッパー 戻; [10] 【Y1209】コンテナ仕分けストッパー 行; [11] 【Y1210】コンテナ仕分け送り 戻 *)
END_VAR
VAR_GLOBAL
    Out_CYw_Hnd_Feed_B_F_Done : BOOL;  (* 【Y1303】B(右側) コンベア受渡送り行 動作完了 *)
    Out_CYw_Hnd_Feed_B_F_Manual : ARRAY[0..10] OF Bool;  (* 手動【Y1303】B(右側) コンベア受渡送り行： *)
    Out_CYw_Hnd_Feed_B_F_Auto : ARRAY[0..10] OF Bool;  (* 自動【Y1303】B(右側) コンベア受渡送り行： *)
    Out_CYw_Hnd_Feed_B_H_Done : BOOL;  (* 【Y1302】B(右側) コンベア受渡送り戻 動作完了 *)
    Out_CYw_Hnd_Feed_B_H_Manual : ARRAY[0..10] OF Bool;  (* 手動【Y1302】B(右側) コンベア受渡送り戻： *)
    Out_CYw_Hnd_Feed_B_H_Auto : ARRAY[0..10] OF Bool;  (* 自動【Y1302】B(右側) コンベア受渡送り戻： *)
    Out_CYw_Hnd_Feed_A_F_Done : BOOL;  (* 【Y1301】A(左側) コンベア受渡送り行 動作完了 *)
    Out_CYw_Hnd_Feed_A_F_Manual : ARRAY[0..10] OF Bool;  (* 手動【Y1301】A(左側) コンベア受渡送り行： *)
    Out_CYw_Srt_Feed_H_Manual : ARRAY[0..10] OF Bool;  (* 手動【Y1210】コンテナ仕分け送り 戻： *)
    Out_CYw_Srt_Feed_H_Done : BOOL;  (* 【Y1210】コンテナ仕分け送り 戻 動作完了 *)
    Out_CYw_Srt_Feed_F_Auto : ARRAY[0..10] OF Bool;  (* 自動【Y1211】コンテナ仕分け送り 行： *)
    Out_CYw_Srt_Feed_F_Manual : ARRAY[0..10] OF Bool;  (* 手動【Y1211】コンテナ仕分け送り 行： *)
    Out_CYw_Srt_Feed_F_Done : BOOL;  (* 【Y1211】コンテナ仕分け送り 行 動作完了 *)
    Out_CYw_Hnd_Feed_A_H_Auto : ARRAY[0..10] OF Bool;  (* 自動【Y1300】A(左側) コンベア受渡送り戻： *)
    Out_CYw_Hnd_Feed_A_H_Manual : ARRAY[0..10] OF Bool;  (* 手動【Y1300】A(左側) コンベア受渡送り戻： *)
    Out_CYw_Hnd_Feed_A_H_Done : BOOL;  (* 【Y1300】A(左側) コンベア受渡送り戻 動作完了 *)
    Out_CYw_Hnd_Feed_A_F_Auto : ARRAY[0..10] OF Bool;  (* 自動【Y1301】A(左側) コンベア受渡送り行： *)
    Out_CYw_Empty_Container_CY_F_Done : BOOL;  (* 【Y1201】空コンテナ送り 行 動作完了 *)
    Out_CYw_Sep_Claw_H_Auto : ARRAY[0..10] OF Bool;  (* 自動【Y1202】段バラシ爪 戻： *)
    Out_CYw_Sep_Claw_H_Manual : ARRAY[0..10] OF Bool;  (* 手動【Y1202】段バラシ爪 戻： *)
    Out_CYw_Sep_Claw_H_Done : BOOL;  (* 【Y1202】段バラシ爪 戻 動作完了 *)
    Out_CYw_Sep_Claw_F_Auto : ARRAY[0..10] OF Bool;  (* 自動【Y1203】段バラシ爪 行： *)
    Out_CYw_Sep_Claw_F_Manual : ARRAY[0..10] OF Bool;  (* 手動【Y1203】段バラシ爪 行： *)
    Out_CYw_Sep_Claw_F_Done : BOOL;  (* 【Y1203】段バラシ爪 行 動作完了 *)
    Out_CYw_Ejc_Cont_H_Auto : ARRAY[0..10] OF Bool;  (* 自動【Y1204】コンテナ排出 戻： *)
    Out_CYw_Ejc_Cont_H_Manual : ARRAY[0..10] OF Bool;  (* 手動【Y1204】コンテナ排出 戻： *)
    Out_CYw_Ejc_Cont_H_Done : BOOL;  (* 【Y1204】コンテナ排出 戻 動作完了 *)
    Out_CYw_Ejc_Cont_F_Auto : ARRAY[0..10] OF Bool;  (* 自動【Y1205】コンテナ排出 行： *)
    Out_CYw_Ejc_Cont_F_Manual : ARRAY[0..10] OF Bool;  (* 手動【Y1205】コンテナ排出 行： *)
    Out_CYw_Ejc_Cont_F_Done : BOOL;  (* 【Y1205】コンテナ排出 行 動作完了 *)
    Out_CYw_Box_Chuck_H_Auto : ARRAY[0..10] OF Bool;  (* 自動【Y1206】箱入れチャック 戻： *)
    Out_CYw_Box_Chuck_H_Manual : ARRAY[0..10] OF Bool;  (* 手動【Y1206】箱入れチャック 戻： *)
    Out_CYw_Box_Chuck_H_Done : BOOL;  (* 【Y1206】箱入れチャック 戻 動作完了 *)
    Out_CYw_Box_Chuck_F_Auto : ARRAY[0..10] OF Bool;  (* 自動【Y1207】箱入れチャック 行： *)
    Out_CYw_Box_Chuck_F_Manual : ARRAY[0..10] OF Bool;  (* 手動【Y1207】箱入れチャック 行： *)
    Out_CYw_Box_Chuck_F_Done : BOOL;  (* 【Y1207】箱入れチャック 行 動作完了 *)
    Out_CYw_Srt_Stopper_H_Auto : ARRAY[0..10] OF Bool;  (* 自動【Y1208】コンテナ仕分けストッパー 戻： *)
    Out_CYw_Srt_Stopper_H_Manual : ARRAY[0..10] OF Bool;  (* 手動【Y1208】コンテナ仕分けストッパー 戻 行： *)
    Out_CYw_Srt_Stopper_H_Done : BOOL;  (* 【Y1208】コンテナ仕分けストッパー 戻 動作完了 *)
    Out_CYw_Srt_Stopper_F_Auto : ARRAY[0..10] OF Bool;  (* 自動【Y1209】コンテナ仕分けストッパー 行： *)
    Out_CYw_Srt_Stopper_F_Manual : ARRAY[0..10] OF Bool;  (* 手動【Y1209】コンテナ仕分けストッパー 行： *)
    Out_CYw_Srt_Stopper_F_Done : BOOL;  (* 【Y1209】コンテナ仕分けストッパー 行 動作完了 *)
    Out_CYw_Srt_Feed_H_Auto : ARRAY[0..10] OF Bool;  (* 自動【Y1210】コンテナ仕分け送り 戻： *)
    Out_CYS_Pos_04_Stopper_B_H_Auto : ARRAY[0..10] OF Bool;  (* 自動【Y823】B(右側) 位置4ストッパー戻： *)
    Out_CYS_Pos_04_Stopper_B_H_Manual : ARRAY[0..10] OF Bool;  (* 手動【Y823】B(右側) 位置4ストッパー戻： *)
    Out_CYS_Pos_04_Stopper_B_H_Done : BOOL;  (* 【Y823】B(右側) 位置4ストッパー戻 動作完了 *)
    Out_CYS_Pos_04_Stopper_B_F_Auto : ARRAY[0..10] OF Bool;  (* 自動【Y823】B(右側) 位置4ストッパー行： *)
    Out_CYS_Pos_04_Stopper_B_F_Manual : ARRAY[0..10] OF Bool;  (* 手動【Y823】B(右側) 位置4ストッパー行： *)
    Out_CYS_Pos_04_Stopper_B_F_Done : BOOL;  (* 【Y823】B(右側) 位置4ストッパー行 動作完了 *)
    Out_CYS_Pos_05_Stopper_B_H_Auto : ARRAY[0..10] OF Bool;  (* 自動【Y824】B(右側) 位置5ストッパー戻： *)
    Out_CYS_Pos_05_Stopper_B_H_Manual : ARRAY[0..10] OF Bool;  (* 手動【Y824】B(右側) 位置5ストッパー戻： *)
    Out_CYS_Pos_05_Stopper_B_H_Done : BOOL;  (* 【Y824】B(右側) 位置5ストッパー戻 動作完了 *)
    Out_CYS_Pos_05_Stopper_B_F_Auto : ARRAY[0..10] OF Bool;  (* 自動【Y824】B(右側) 位置5ストッパー行： *)
    Out_CYS_Pos_05_Stopper_B_F_Manual : ARRAY[0..10] OF Bool;  (* 手動【Y824】B(右側) 位置5ストッパー行： *)
    Out_CYS_Pos_05_Stopper_B_F_Done : BOOL;  (* 【Y824】B(右側) 位置5ストッパー行 動作完了 *)
    Out_CYS_Pos_06_Stopper_B_H_Auto : ARRAY[0..10] OF Bool;  (* 自動【Y825】B(右側) 位置6ストッパー戻： *)
    Out_CYS_Pos_06_Stopper_B_H_Manual : ARRAY[0..10] OF Bool;  (* 手動【Y825】B(右側) 位置6ストッパー戻： *)
    Out_CYS_Pos_06_Stopper_B_H_Done : BOOL;  (* 【Y825】B(右側) 位置6ストッパー戻 動作完了 *)
    Out_CYS_Pos_06_Stopper_B_F_Auto : ARRAY[0..10] OF Bool;  (* 自動【Y825】B(右側) 位置6ストッパー行： *)
    Out_CYS_Pos_06_Stopper_B_F_Manual : ARRAY[0..10] OF Bool;  (* 手動【Y825】B(右側) 位置6ストッパー行： *)
    Out_CYS_Pos_06_Stopper_B_F_Done : BOOL;  (* 【Y825】B(右側) 位置6ストッパー行 動作完了 *)
    Out_CYw_SH_B_Turn_H_Auto : ARRAY[0..10] OF Bool;  (* 自動【Y826】B(右側) ストックフォルダターン戻： *)
    Out_CYw_SH_B_Turn_H_Manual : ARRAY[0..10] OF Bool;  (* 手動【Y826】B(右側) ストックフォルダターン戻： *)
    Out_CYw_SH_B_Turn_H_Done : BOOL;  (* 【Y826】B(右側) ストックフォルダターン戻 動作完了 *)
    Out_CYw_SH_B_Turn_F_Manual : ARRAY[0..10] OF Bool;  (* 自動【Y827】B(右側) ストックフォルダターン行： *)
    Out_CYw_SH_B_Turn_F_Auto : ARRAY[0..10] OF Bool;  (* 手動【Y827】B(右側) ストックフォルダターン行： *)
    Out_CYw_SH_B_Turn_F_Done : BOOL;  (* 【Y827】B(右側) ストックフォルダターン行 動作完了 *)
    Out_CYw_NG1_Srt_B_H_Auto : ARRAY[0..10] OF Bool;  (* 自動【Y828】B(右側) NG1仕分け 戻： *)
    Out_CYw_NG1_Srt_B_H_Manual : ARRAY[0..10] OF Bool;  (* 手動【Y828】B(右側) NG1仕分け 戻： *)
    Out_CYw_NG1_Srt_B_H_Done : BOOL;  (* 【Y828】B(右側) NG1仕分け 戻 動作完了 *)
    Out_CYw_NG1_Srt_B_F_Auto : ARRAY[0..10] OF Bool;  (* 自動【Y829】B(右側) NG1仕分け 行： *)
    Out_CYw_NG1_Srt_B_F_Manual : ARRAY[0..10] OF Bool;  (* 手動【Y829】B(右側) NG1仕分け 行： *)
    Out_CYw_NG1_Srt_B_F_Done : BOOL;  (* 【Y829】B(右側) NG1仕分け 行 動作完了 *)
    Out_CYw_Empty_Container_CY_H_Manual : ARRAY[0..10] OF Bool;  (* 手動【Y1200】空コンテナ送り 戻： *)
    Out_CYw_Empty_Container_CY_H_Auto : ARRAY[0..10] OF Bool;  (* 自動【Y1200】空コンテナ送り 戻： *)
    Out_CYw_Empty_Container_CY_H_Done : BOOL;  (* 【Y1200】空コンテナ送り 戻 動作完了 *)
    Out_CYw_Empty_Container_CY_F_Auto : ARRAY[0..10] OF Bool;  (* 自動【Y1201】空コンテナ送り 行： *)
    Out_CYw_Empty_Container_CY_F_Manual : ARRAY[0..10] OF Bool;  (* 手動【Y1201】空コンテナ送り 行： *)
    Out_CYw_Rev_02_Pick_B_H_Manual : ARRAY[0..10] OF Bool;  (* 手動【Y814】B(右側)ST6 反転2ピックアップ戻： *)
    Out_CYw_Rev_02_Pick_B_H_Done : BOOL;  (* 【Y814】B(右側)ST6 反転2ピックアップ戻 動作完了 *)
    Out_CYw_Rev_02_Pick_B_F_Auto : ARRAY[0..10] OF Bool;  (* 自動【Y815】B(右側)ST6 反転2ピックアップ行 ： *)
    Out_CYw_Rev_02_Pick_B_F_Manual : ARRAY[0..10] OF Bool;  (* 手動【Y815】B(右側)ST6 反転2ピックアップ行： *)
    Out_CYw_Rev_02_Pick_B_F_Done : BOOL;  (* 【Y815】B(右側)ST6 反転2ピックアップ行 動作完了 *)
    Out_CYw_Disc_Chk_B_H_Auto : ARRAY[0..10] OF Bool;  (* 自動【Y816】B(右側) 排出チャック閉 戻 ： *)
    Out_CYw_Disc_Chk_B_H_Manual : ARRAY[0..10] OF Bool;  (* 手動【Y816】B(右側) 排出チャック閉 戻： *)
    Out_CYw_Disc_Chk_B_H_Done : BOOL;  (* 【Y816】B(右側) 排出チャック閉 戻 動作完了 *)
    Out_CYw_Disc_Chk_B_F_Auto : ARRAY[0..10] OF Bool;  (* 自動【Y817】B(右側) 排出チャック開 行 ： *)
    Out_CYw_Disc_Chk_B_F_Manual : ARRAY[0..10] OF Bool;  (* 手動【Y817】B(右側) 排出チャック開 行： *)
    Out_CYw_Disc_Chk_B_F_Done : BOOL;  (* 【Y817】B(右側) 排出チャック開 行 動作完了 *)
    Out_CYw_Ejc_Hldr_Feed_B_H_Auto : ARRAY[0..10] OF Bool;  (* 自動【Y818】B(右側) 排出フォルダ送り戻： *)
    Out_CYw_Ejc_Hldr_Feed_B_H_Manual : ARRAY[0..10] OF Bool;  (* 手動【Y818】B(右側) 排出フォルダ送り戻： *)
    Out_CYw_Ejc_Hldr_Feed_B_H_Done : BOOL;  (* 【Y818】B(右側) 排出フォルダ送り戻 動作完了 *)
    Out_CYw_Ejc_Hldr_Feed_B_F_Auto : ARRAY[0..10] OF Bool;  (* 自動【Y819】B(右側) 排出フォルダ送り行： *)
    Out_CYw_Ejc_Hldr_Feed_B_F_Manual : ARRAY[0..10] OF Bool;  (* 手動【Y819】B(右側) 排出フォルダ送り行： *)
    Out_CYw_Ejc_Hldr_Feed_B_F_Done : BOOL;  (* 【Y819】B(右側) 排出フォルダ送り行 動作完了 *)
    Out_CYS_Pos_01_Stopper_B_H_Auto : ARRAY[0..10] OF Bool;  (* 自動【Y820】B(右側) 位置1ストッパー戻： *)
    Out_CYS_Pos_01_Stopper_B_H_Manual : ARRAY[0..10] OF Bool;  (* 手動【Y820】B(右側) 位置1ストッパー戻： *)
    Out_CYS_Pos_01_Stopper_B_H_Done : BOOL;  (* 【Y820】B(右側) 位置1ストッパー戻 動作完了 *)
    Out_CYS_Pos_01_Stopper_B_F_Auto : ARRAY[0..10] OF Bool;  (* 自動【Y820】B(右側) 位置1ストッパー 行： *)
    Out_CYS_Pos_01_Stopper_B_F_Manual : ARRAY[0..10] OF Bool;  (* 手動【Y820】B(右側) 位置1ストッパー 行： *)
    Out_CYS_Pos_01_Stopper_B_F_Done : BOOL;  (* 【Y820】B(右側) 位置1ストッパー 行 動作完了 *)
    Out_CYS_Pos_02_Stopper_B_H_Auto : ARRAY[0..10] OF Bool;  (* 自動【Y821】B(右側) 位置2ストッパー戻： *)
    Out_CYS_Pos_02_Stopper_B_H_Manual : ARRAY[0..10] OF Bool;  (* 手動【Y821】B(右側) 位置2ストッパー戻： *)
    Out_CYS_Pos_02_Stopper_B_H_Done : BOOL;  (* 【Y821】B(右側) 位置2ストッパー戻 動作完了 *)
    Out_CYS_Pos_02_Stopper_B_F_Auto : ARRAY[0..10] OF Bool;  (* 自動【Y821】B(右側) 位置2ストッパー行： *)
    Out_CYS_Pos_02_Stopper_B_F_Manual : ARRAY[0..10] OF Bool;  (* 手動【Y821】B(右側) 位置2ストッパー行： *)
    Out_CYS_Pos_02_Stopper_B_F_Done : BOOL;  (* 【Y821】B(右側) 位置2ストッパー行 動作完了 *)
    Out_CYS_Pos_03_Stopper_B_H_Auto : ARRAY[0..10] OF Bool;  (* 自動【Y822】B(右側) 位置3ストッパー戻： *)
    Out_CYS_Pos_03_Stopper_B_H_Manual : ARRAY[0..10] OF Bool;  (* 手動【Y822】B(右側) 位置3ストッパー戻： *)
    Out_CYS_Pos_03_Stopper_B_H_Done : BOOL;  (* 【Y822】B(右側) 位置3ストッパー戻 動作完了 *)
    Out_CYS_Pos_03_Stopper_B_F_Auto : ARRAY[0..10] OF Bool;  (* 自動【Y822】B(右側) 位置3ストッパー行： *)
    Out_CYS_Pos_03_Stopper_B_F_Manual : ARRAY[0..10] OF Bool;  (* 手動【Y822】B(右側) 位置3ストッパー行： *)
    Out_CYS_Pos_03_Stopper_B_F_Done : BOOL;  (* 【Y822】B(右側) 位置3ストッパー行 動作完了 *)
    Out_CYw_HgtInsp_Lf_B_H_Done : BOOL;  (* 【Y802】B(右側) 高さ検査持上戻 動作完了 *)
    Out_CYw_HgtInsp_Lf_B_F_Auto : ARRAY[0..10] OF Bool;  (* 自動【Y803】B(右側) 高さ検査持上行： *)
    Out_CYw_HgtInsp_Lf_B_F_Manual : ARRAY[0..10] OF Bool;  (* 手動【Y803】B(右側) 高さ検査持上行： *)
    Out_CYw_HgtInsp_Lf_B_F_Done : BOOL;  (* 【Y803】B(右側) 高さ検査持上行 動作完了 *)
    Out_CYw_NG1_Pick_B_H_Auto : ARRAY[0..10] OF Bool;  (* 自動【Y804】B(右側) NG1ピックアップ戻： *)
    Out_CYw_NG1_Pick_B_H_Manual : ARRAY[0..10] OF Bool;  (* 手動【Y804】B(右側) NG1ピックアップ戻： *)
    Out_CYw_NG1_Pick_B_H_Done : BOOL;  (* 【Y804】B(右側) NG1ピックアップ戻 動作完了 *)
    Out_CYw_NG1_Pick_B_F_Auto : ARRAY[0..10] OF Bool;  (* 自動【Y805】B(右側) NG1ピックアップ行： *)
    Out_CYw_NG1_Pick_B_F_Manual : ARRAY[0..10] OF Bool;  (* 手動【Y805】B(右側) NG1ピックアップ行： *)
    Out_CYw_NG1_Pick_B_F_Done : BOOL;  (* 【Y805】B(右側) NG1ピックアップ行 動作完了 *)
    Out_CYw_NG1_Chk_B_H_Auto : ARRAY[0..10] OF Bool;  (* 自動【Y806】B(右側) NG1チャック戻： *)
    Out_CYw_NG1_Chk_B_H_Manual : ARRAY[0..10] OF Bool;  (* 手動【Y806】B(右側) NG1チャック戻： *)
    Out_CYw_NG1_Chk_B_H_Done : BOOL;  (* 【Y806】B(右側) NG1チャック戻 動作完了 *)
    Out_CYw_NG1_Chk_B_F_Auto : ARRAY[0..10] OF Bool;  (* 自動【Y807】B(右側) NG1チャック行： *)
    Out_CYw_NG1_Chk_B_F_Manual : ARRAY[0..10] OF Bool;  (* 手動【Y807】B(右側) NG1チャック行： *)
    Out_CYw_NG1_Chk_B_F_Done : BOOL;  (* 【Y807】B(右側) NG1チャック行 動作完了 *)
    Out_CYw_Rev_01_Chk_B_H_Auto : ARRAY[0..10] OF Bool;  (* 自動【Y808】B(右側)ST4 反転1チャック閉 戻： *)
    Out_CYw_Rev_01_Chk_B_H_Manual : ARRAY[0..10] OF Bool;  (* 手動【Y808】B(右側)ST4 反転1チャック閉 戻： *)
    Out_CYw_Rev_01_Chk_B_H_Done : BOOL;  (* 【Y808】B(右側)ST4 反転1チャック閉 戻 動作完了 *)
    Out_CYw_Rev_01_Chk_B_F_Auto : ARRAY[0..10] OF Bool;  (* 自動【Y809】B(右側)ST4 反転1チャック開 戻： *)
    Out_CYw_Rev_01_Chk_B_F_Manual : ARRAY[0..10] OF Bool;  (* 手動【Y809】B(右側)ST4 反転1チャック開 戻： *)
    Out_CYw_Rev_01_Chk_B_F_Done : BOOL;  (* 【Y809】B(右側)ST4 反転1チャック開 戻 動作完了 *)
    Out_CYw_Rev_01_Pick_B_H_Auto : ARRAY[0..10] OF Bool;  (* 自動【Y810】B(右側)ST4 反転1ピックアップ戻： *)
    Out_CYw_Rev_01_Pick_B_H_Manual : ARRAY[0..10] OF Bool;  (* 手動【Y810】B(右側)ST4 反転1ピックアップ戻： *)
    Out_CYw_Rev_01_Pick_B_H_Done : BOOL;  (* 【Y810】B(右側)ST4 反転1ピックアップ戻 動作完了 *)
    Out_CYw_Rev_01_Pick_B_F_Auto : ARRAY[0..10] OF Bool;  (* 自動【Y811】B(右側)ST4 反転1ピックアップ行： *)
    Out_CYw_Rev_01_Pick_B_F_Manual : ARRAY[0..10] OF Bool;  (* 手動【Y811】B(右側)ST4 反転1ピックアップ行： *)
    Out_CYw_Rev_01_Pick_B_F_Done : BOOL;  (* 【Y811】B(右側)ST4 反転1ピックアップ行 動作完了 *)
    Out_CYw_Rev_02_Chk_B_H_Auto : ARRAY[0..10] OF Bool;  (* 自動【Y812】B(右側)ST6 反転2チャック閉 戻： *)
    Out_CYw_Rev_02_Chk_B_H_Manual : ARRAY[0..10] OF Bool;  (* 手動【Y812】B(右側)ST6 反転2チャック閉 戻： *)
    Out_CYw_Rev_02_Chk_B_H_Done : BOOL;  (* 【Y812】B(右側)ST6 反転2チャック閉 戻 動作完了 *)
    Out_CYw_Rev_02_Chk_B_F_Auto : ARRAY[0..10] OF Bool;  (* 自動【Y813】B(右側)ST6 反転2チャック開 行 ： *)
    Out_CYw_Rev_02_Chk_B_F_Manual : ARRAY[0..10] OF Bool;  (* 手動【Y813】B(右側)ST6 反転2チャック開 行： *)
    Out_CYw_Rev_02_Chk_B_F_Done : BOOL;  (* 【Y813】B(右側)ST6 反転2チャック開 行 動作完了 *)
    Out_CYw_Rev_02_Pick_B_H_Auto : ARRAY[0..10] OF Bool;  (* 自動【Y814】B(右側)ST6 反転2ピックアップ戻 ： *)
    Out_CYw_HgtInsp_Clp_B_H_Done : BOOL;  (* 【Y800】B(右側) 高さ検査押え戻 動作完了 *)
    Out_CYw_HgtInsp_Clp_B_H_Auto : ARRAY[0..10] OF Bool;  (* 自動【Y800】B(右側) 高さ検査押え戻： *)
    Out_CYw_HgtInsp_Clp_B_H_Manual : ARRAY[0..10] OF Bool;  (* 手動【Y800】B(右側) 高さ検査押え戻： *)
    Out_CYw_HgtInsp_Clp_B_F_Auto : ARRAY[0..10] OF Bool;  (* 自動【Y801】B(右側) 高さ検査押え行： *)
    Out_CYw_HgtInsp_Clp_B_F_Manual : ARRAY[0..10] OF Bool;  (* 手動【Y801】B(右側) 高さ検査押え行： *)
    Out_CYw_HgtInsp_Clp_B_F_Done : BOOL;  (* 【Y801】B(右側) 高さ検査押え行 動作完了 *)
    Out_CYw_HgtInsp_Lf_B_H_Auto : ARRAY[0..10] OF Bool;  (* 自動【Y802】B(右側) 高さ検査持上戻： *)
    Out_CYw_HgtInsp_Lf_B_H_Manual : ARRAY[0..10] OF Bool;  (* 手動【Y802】B(右側) 高さ検査持上戻： *)
    Out_CYS_Pos_03_Stopper_A_H_Manual : ARRAY[0..10] OF Bool;  (* 手動【Y722】A(左側) 位置3ストッパー戻： *)
    Out_CYS_Pos_03_Stopper_A_H_Done : BOOL;  (* 【Y722】A(左側) 位置3ストッパー戻 動作完了 *)
    Out_CYS_Pos_03_Stopper_A_F_Auto : ARRAY[0..10] OF Bool;  (* 自動【Y722】A(左側) 位置3ストッパー行： *)
    Out_CYS_Pos_03_Stopper_A_F_Manual : ARRAY[0..10] OF Bool;  (* 手動【Y722】A(左側) 位置3ストッパー行： *)
    Out_CYS_Pos_03_Stopper_A_F_Done : BOOL;  (* 【Y722】A(左側) 位置3ストッパー行 動作完了 *)
    Out_CYS_Pos_04_Stopper_A_H_Auto : ARRAY[0..10] OF Bool;  (* 自動【Y723】A(左側) 位置4ストッパー戻：; [1] A(左側)検査完了後; [2] A(左側)原点位置移動 *)
    Out_CYS_Pos_04_Stopper_A_H_Manual : ARRAY[0..10] OF Bool;  (* 手動【Y723】A(左側) 位置4ストッパー戻： *)
    Out_CYS_Pos_04_Stopper_A_H_Done : BOOL;  (* 【Y723】A(左側) 位置4ストッパー戻 動作完了 *)
    Out_CYS_Pos_04_Stopper_A_F_Auto : ARRAY[0..10] OF Bool;  (* 自動【Y723】A(左側) 位置4ストッパー行： *)
    Out_CYS_Pos_04_Stopper_A_F_Manual : ARRAY[0..10] OF Bool;  (* 手動【Y723】A(左側) 位置4ストッパー行： *)
    Out_CYS_Pos_04_Stopper_A_F_Done : BOOL;  (* 【Y723】A(左側) 位置4ストッパー行 動作完了 *)
    Out_CYS_Pos_05_Stopper_A_H_Auto : ARRAY[0..10] OF Bool;  (* 自動【Y724】A(左側) 位置5ストッパー戻：; [1] A(左側)検査完了後; [2] A(左側) ST5 カメラ2検査開始 *)
    Out_CYS_Pos_05_Stopper_A_H_Manual : ARRAY[0..10] OF Bool;  (* 手動【Y724】A(左側) 位置5ストッパー戻： *)
    Out_CYS_Pos_05_Stopper_A_H_Done : BOOL;  (* 【Y724】A(左側) 位置5ストッパー戻 動作完了 *)
    Out_CYS_Pos_05_Stopper_A_F_Auto : ARRAY[0..10] OF Bool;  (* 自動【Y724】A(左側) 位置5ストッパー行： *)
    Out_CYS_Pos_05_Stopper_A_F_Manual : ARRAY[0..10] OF Bool;  (* 手動【Y724】A(左側) 位置5ストッパー行： *)
    Out_CYS_Pos_05_Stopper_A_F_Done : BOOL;  (* 【Y724】A(左側) 位置5ストッパー行 動作完了 *)
    Out_CYS_Pos_06_Stopper_A_H_Auto : ARRAY[0..10] OF Bool;  (* 自動【Y725】A(左側) 位置6ストッパー戻：; [1] A(左側)検査完了後; [2] A(左側) ST6 原点位置移動 *)
    Out_CYS_Pos_06_Stopper_A_H_Manual : ARRAY[0..10] OF Bool;  (* 手動【Y725】A(左側) 位置6ストッパー戻： *)
    Out_CYS_Pos_06_Stopper_A_H_Done : BOOL;  (* 【Y725】A(左側) 位置6ストッパー戻 動作完了 *)
    Out_CYS_Pos_06_Stopper_A_F_Auto : ARRAY[0..10] OF Bool;  (* 自動【Y725】A(左側) 位置6ストッパー行： *)
    Out_CYS_Pos_06_Stopper_A_F_Manual : ARRAY[0..10] OF Bool;  (* 手動【Y725】A(左側) 位置6ストッパー行： *)
    Out_CYS_Pos_06_Stopper_A_F_Done : BOOL;  (* 【Y725】A(左側) 位置6ストッパー行 動作完了 *)
    Out_CYw_SH_A_Turn_H_Auto : ARRAY[0..10] OF Bool;  (* 自動【Y726】A(左側) ストックフォルダターン戻： *)
    Out_CYw_SH_A_Turn_H_Manual : ARRAY[0..10] OF Bool;  (* 手動【Y726】A(左側) ストックフォルダターン戻： *)
    Out_CYw_SH_A_Turn_H_Done : BOOL;  (* 【Y726】A(左側) ストックフォルダターン戻 動作完了 *)
    Out_CYw_SH_A_Turn_F_Auto : ARRAY[0..10] OF Bool;  (* 自動【Y727】A(左側) ストックフォルダターン行： *)
    Out_CYw_SH_A_Turn_F_Manual : ARRAY[0..10] OF Bool;  (* 手動【Y727】A(左側) ストックフォルダターン行： *)
    Out_CYw_SH_A_Turn_F_Done : BOOL;  (* 【Y727】A(左側) ストックフォルダターン行 動作完了 *)
    Out_CYw_NG1_Srt_A_H_Auto : ARRAY[0..10] OF Bool;  (* 自動【Y728】A(左側) NG1仕分け 戻：; [1] A(左側)原点位置移動; [2] NGワーク分離 *)
    Out_CYw_NG1_Srt_A_H_Manual : ARRAY[0..10] OF Bool;  (* 手動【Y728】A(左側) NG1仕分け 戻： *)
    Out_CYw_NG1_Srt_A_H_Done : BOOL;  (* 【Y728】A(左側) NG1仕分け 戻 動作完了 *)
    Out_CYw_NG1_Srt_A_F_Auto : ARRAY[0..10] OF Bool;  (* 自動【Y729】A(左側) NG1仕分け行：; [1] NGワーク分離 *)
    Out_CYw_NG1_Srt_A_F_Manual : ARRAY[0..10] OF Bool;  (* 手動【Y729】A(左側) NG1仕分け行： *)
    Out_CYw_NG1_Srt_A_F_Done : BOOL;  (* 【Y729】A(左側) NG1仕分け行 動作完了 *)
    Out_CYS_Pos_01_Stopper_A_F_Auto : ARRAY[0..10] OF Bool;  (* 自動【Y720】A(左側) 位置1ストッパー行： *)
    Out_CYS_Pos_01_Stopper_A_F_Manual : ARRAY[0..10] OF Bool;  (* 手動【Y720】A(左側) 位置1ストッパー 行： *)
    Out_CYS_Pos_02_Stopper_A_H_Auto : ARRAY[0..10] OF Bool;  (* 自動【Y721】A(左側) 位置2ストッパー戻：; [1] A(左側)検査完了後; [2] 原点位置移動 *)
    Out_CYS_Pos_02_Stopper_A_H_Manual : ARRAY[0..10] OF Bool;  (* 手動【Y721】A(左側) 位置2ストッパー戻： *)
    Out_CYS_Pos_02_Stopper_A_H_Done : BOOL;  (* 【Y721】A(左側) 位置2ストッパー戻 動作完了 *)
    Out_CYS_Pos_02_Stopper_A_F_Auto : ARRAY[0..10] OF Bool;  (* 自動【Y721】A(左側) 位置2ストッパー行： *)
    Out_CYS_Pos_02_Stopper_A_F_Manual : ARRAY[0..10] OF Bool;  (* 手動【Y721】A(左側) 位置2ストッパー行： *)
    Out_CYS_Pos_02_Stopper_A_F_Done : BOOL;  (* 【Y721】A(左側) 位置2ストッパー行 動作完了 *)
    Out_CYS_Pos_03_Stopper_A_H_Auto : ARRAY[0..10] OF Bool;  (* 自動【Y722】A(左側) 位置3ストッパー戻：; [1] A(左側)検査完了後; [2] A(左側)原点位置移動 *)
    Out_CYw_Rev_02_Pick_A_H_Auto : ARRAY[0..10] OF Bool;  (* 自動【Y714】A(左側)ST6 反転2ピックアップ戻 ：; [1] A(左側) ST6 反転前戻; [2] A(左側) ST6 設置後戻 *)
    Out_CYw_Rev_02_Pick_A_H_Manual : ARRAY[0..10] OF Bool;  (* 手動【Y714】A(左側)ST6 反転2ピックアップ戻 ： *)
    Out_CYw_Rev_02_Pick_A_H_Done : BOOL;  (* 【Y714】A(左側)ST6 反転2ピックアップ戻 動作完了 *)
    Out_CYw_Rev_02_Pick_A_F_Auto : ARRAY[0..10] OF Bool;  (* 自動【Y715】A(左側)ST6 反転2ピックアップ行 ：; [1] A(左側) ST6 反転前行; [2] A(左側) ST6 設置行 *)
    Out_CYw_Rev_02_Pick_A_F_Manual : ARRAY[0..10] OF Bool;  (* 手動【Y715】A(左側)ST6 反転2ピックアップ行 ： *)
    Out_CYw_Rev_02_Pick_A_F_Done : BOOL;  (* 【Y715】A(左側)ST6 反転2ピックアップ行 動作完了 *)
    Out_CYw_Disc_Chk_A_H_Auto : ARRAY[0..10] OF Bool;  (* 自動【Y716】A(左側) 排出チャック閉 戻 ： *)
    Out_CYw_Disc_Chk_A_H_Manual : ARRAY[0..10] OF Bool;  (* 手動【Y716】A(左側) 排出チャック閉 戻 ： *)
    Out_CYw_Disc_Chk_A_H_Done : BOOL;  (* 【Y716】A(左側) 排出チャック閉 戻 動作完了 *)
    Out_CYw_Disc_Chk_A_F_Auto : ARRAY[0..10] OF Bool;  (* 自動【Y717】A(左側) 排出チャック開 行 ： *)
    Out_CYw_Disc_Chk_A_F_Manual : ARRAY[0..10] OF Bool;  (* 手動【Y717】A(左側) 排出チャック開 行 ： *)
    Out_CYw_Disc_Chk_A_F_Done : BOOL;  (* 【Y717】A(左側) 排出チャック開 行 動作完了 *)
    Out_CYw_Ejc_Hldr_Feed_A_F_Auto : ARRAY[0..10] OF Bool;  (* 自動【Y719】A(左側) 排出フォルダ送り行 ： *)
    Out_CYw_Ejc_Hldr_Feed_A_F_Manual : ARRAY[0..10] OF Bool;  (* 手動【Y719】A(左側) 排出フォルダ送り行 ： *)
    Out_CYw_Ejc_Hldr_Feed_A_F_Done : BOOL;  (* 【Y719】A(左側) 排出フォルダ送り行 動作完了 *)
    Out_CYw_Ejc_Hldr_Feed_A_H_Auto : ARRAY[0..10] OF Bool;  (* 自動【Y718】A(左側) 排出フォルダ送り戻 ： *)
    Out_CYw_Ejc_Hldr_Feed_A_H_Manual : ARRAY[0..10] OF Bool;  (* 手動【Y718】A(左側) 排出フォルダ送り戻 ： *)
    Out_CYw_Ejc_Hldr_Feed_A_H_Done : BOOL;  (* 【Y718】A(左側) 排出フォルダ送り戻 動作完了 *)
    Out_CYS_Pos_01_Stopper_A_H_Auto : ARRAY[0..10] OF Bool;  (* 自動【Y720】A(左側) 位置1ストッパー 戻：; [1] A(左側)検査完了後; [2] 検査開始 *)
    Out_CYS_Pos_01_Stopper_A_H_Manual : ARRAY[0..10] OF Bool;  (* 手動【Y720】A(左側) 位置1ストッパー 戻 ： *)
    Out_CYS_Pos_01_Stopper_A_F_Done : BOOL;  (* 【Y720】A(左側) 位置1ストッパー行 動作完了 *)
    Out_CYS_Pos_01_Stopper_A_H_Done : BOOL;  (* 【Y720】A(左側) 位置1ストッパー戻 動作完了 *)
    Out_CYw_HgtInsp_Lf_A_F_Done : BOOL;  (* 【Y703】A(左側) 高さ検査持上行 動作完了 *)
    Out_CYw_NG1_Pick_A_H_Auto : ARRAY[0..10] OF Bool;  (* 自動【Y704】A(左側) NG1ピックアップ戻：; [1] A(左側)原点位置移動; [2] NGワーク回収 *)
    Out_CYw_NG1_Pick_A_H_Manual : ARRAY[0..10] OF Bool;  (* 手動【Y704】A(左側) NG1ピックアップ戻： *)
    Out_CYw_NG1_Pick_A_H_Done : BOOL;  (* 【Y704】A(左側) NG1ピックアップ戻 動作完了 *)
    Out_CYw_NG1_Pick_A_F_Auto : ARRAY[0..10] OF Bool;  (* 自動【Y705】A(左側) NG1ピックアップ 行：; [1] NGワーク回収; [2] NG1ワーク切り離し *)
    Out_CYw_NG1_Pick_A_F_Manual : ARRAY[0..10] OF Bool;  (* 手動【Y705】A(左側) NG1ピックアップ 行： *)
    Out_CYw_NG1_Pick_A_F_Done : BOOL;  (* 【Y705】A(左側) NG1ピックアップ 動作完了 *)
    Out_CYw_NG1_Chk_A_H_Auto : ARRAY[0..10] OF Bool;  (* 自動【Y706】A(左側) NG1チャック戻 ：; [1] A(左側)原点位置移動; [2] NGワーク分離 *)
    Out_CYw_NG1_Chk_A_H_Manual : ARRAY[0..10] OF Bool;  (* 手動【Y706】A(左側) NG1チャック戻 ： *)
    Out_CYw_NG1_Chk_A_H_Done : BOOL;  (* 【Y706】A(左側) NG1チャック戻 動作完了 *)
    Out_CYw_NG1_Chk_A_F_Auto : ARRAY[0..10] OF Bool;  (* 自動【Y707】A(左側) NG1チャック行：; [1] NGワーク回収 *)
    Out_CYw_NG1_Chk_A_F_Manual : ARRAY[0..10] OF Bool;  (* 手動【Y707】A(左側) NG1チャック行： *)
    Out_CYw_NG1_Chk_A_F_Done : BOOL;  (* 【Y707】A(左側) NG1チャック行 動作完了 *)
    Out_CYw_Rev_01_Chk_A_H_Auto : ARRAY[0..10] OF Bool;  (* 自動【Y708】A(左側)ST4 反転1チャック閉： *)
    Out_CYw_Rev_01_Chk_A_H_Manual : ARRAY[0..10] OF Bool;  (* 手動【Y708】A(左側)ST4 反転1チャック閉： *)
    Out_CYw_Rev_01_Chk_A_H_Done : BOOL;  (* 【Y708】A(左側)ST4 反転1チャック閉 動作完了 *)
    Mtr_Flip_01_Busy : BOOL;  (* A(左側)反転 オリエンタルモータ1 動作中 *)
    Out_CYw_Rev_01_Chk_A_F_Auto : ARRAY[0..10] OF Bool;  (* 自動【Y709】A(左側)ST4 反転1チャック開： *)
    Out_CYw_Rev_01_Chk_A_F_Manual : ARRAY[0..10] OF Bool;  (* 手動【Y709】A(左側)ST4 反転1チャック開： *)
    Out_CYw_Rev_01_Chk_A_F_Done : BOOL;  (* 【Y709】A(左側)ST4 反転1チャック開 動作完了 *)
    Out_CYw_Rev_01_Pick_A_H_Auto : ARRAY[0..10] OF Bool;  (* 自動【Y710】A(左側)ST4 反転1ピックアップ戻：; [1] ワーク反転動作; [2] 反転後ワーク設置動作 *)
    Out_CYw_Rev_01_Pick_A_H_Manual : ARRAY[0..10] OF Bool;  (* 手動【Y710】A(左側)ST4 反転1ピックアップ戻： *)
    Out_CYw_Rev_01_Pick_A_H_Done : BOOL;  (* 【Y710】A(左側)ST4 反転1ピックアップ戻 動作完了 *)
    Out_CYw_Rev_01_Pick_A_F_Auto : ARRAY[0..10] OF Bool;  (* 自動【Y711】A(左側)ST4 反転1ピックアップ行：; [1] ワーク反転動作; [2] 反転後ワーク設置動作 *)
    Out_CYw_Rev_01_Pick_A_F_Manual : ARRAY[0..10] OF Bool;  (* 手動【Y711】A(左側)ST4 反転1ピックアップ行： *)
    Out_CYw_Rev_01_Pick_A_F_Done : BOOL;  (* 【Y711】A(左側)ST4 反転1ピックアップ行 動作完了 *)
    Out_CYw_Rev_02_Chk_A_H_Auto : ARRAY[0..10] OF Bool;  (* 自動【Y712】A(左側)ST6 反転2チャック閉 戻：; [1] ワーク反転動作 *)
    Out_CYw_Rev_02_Chk_A_H_Manual : ARRAY[0..10] OF Bool;  (* 手動【Y712】A(左側)ST6 反転2チャック閉 戻： *)
    Out_CYw_Rev_02_Chk_A_H_Done : BOOL;  (* 【Y712】A(左側)ST6 反転2チャック閉 戻 動作完了 *)
    Out_CYw_Rev_02_Chk_A_F_Auto : ARRAY[0..10] OF Bool;  (* 自動【Y713】A(左側)ST6 反転2チャック開 行 戻：; [2] 反転後ワーク設置動作; [1] 反転後ワーク設置動作 *)
    Out_CYw_Rev_02_Chk_A_F_Manual : ARRAY[0..10] OF Bool;  (* 手動【Y713】A(左側)ST6 反転2チャック開 行 戻： *)
    Out_CYw_Rev_02_Chk_A_F_Done : BOOL;  (* 【Y713】A(左側)ST6 反転2チャック開 行 動作完了 *)
    Out_CYw_Sply_Slide_B_F_Done : BOOL;  (* 【Y623】B(右側) 供給スライド行 動作完了 *)
    Out_CYw_Sply_Pick_B_H_Auto : ARRAY[0..10] OF Bool;  (* 自動【Y624】B(右側) 供給ピックアップ戻： *)
    Out_CYw_Sply_Pick_B_H_Manual : ARRAY[0..10] OF Bool;  (* 手動【Y624】B(右側) 供給ピックアップ戻： *)
    Out_CYw_Sply_Pick_B_H_Done : BOOL;  (* 【Y624】B(右側) 供給ピックアップ戻 動作完了 *)
    Out_CYw_Sply_Pick_B_F_Auto : ARRAY[0..10] OF Bool;  (* 自動【Y625】B(右側) 供給ピックアップ行： *)
    Out_CYw_Sply_Pick_B_F_Manual : ARRAY[0..10] OF Bool;  (* 手動【Y625】B(右側) 供給ピックアップ行： *)
    Out_CYw_Sply_Pick_B_F_Done : BOOL;  (* 【Y625】B(右側) 供給ピックアップ行 動作完了 *)
    Out_CYw_Sup_Chuck_B_Cl_H_Auto : ARRAY[0..10] OF Bool;  (* 自動【Y626】B(右側) 供給チャック閉 戻： *)
    Out_CYw_Sup_Chuck_B_Cl_H_Manual : ARRAY[0..10] OF Bool;  (* 手動【Y626】B(右側) 供給チャック閉 戻： *)
    Out_CYw_Sup_Chuck_B_Cl_H_Done : BOOL;  (* 【Y626】B(右側) 供給チャック閉 戻 動作完了 *)
    Out_CYw_Sup_Chuck_B_Cl_F_Auto : ARRAY[0..10] OF Bool;  (* 自動【Y627】B(右側) 供給チャック開 行： *)
    Out_CYw_Sup_Chuck_B_Cl_F_Manual : ARRAY[0..10] OF Bool;  (* 手動【Y627】B(右側) 供給チャック開 行： *)
    Out_CYw_Sup_Chuck_B_Cl_F_Done : BOOL;  (* 【Y627】B(右側) 供給チャック開 行 動作完了 *)
    Out_CYw_HgtInsp_Clp_A_H_Auto : ARRAY[0..10] OF Bool;  (* 自動【Y700】A(左側) 高さ検査押え戻：; [1] 原点位置移動 *)
    Out_CYw_HgtInsp_Clp_A_H_Manual : ARRAY[0..10] OF Bool;  (* 手動【Y700】A(左側) 高さ検査押え戻： *)
    Out_CYw_HgtInsp_Clp_A_H_Done : BOOL;  (* 【Y700】A(左側) 高さ検査押え戻 動作完了 *)
    Out_CYw_HgtInsp_Clp_A_F_Auto : ARRAY[0..10] OF Bool;  (* 自動【Y701】A(左側) 高さ検査押え行：; [1] 高さ検査位置 *)
    Out_CYw_HgtInsp_Clp_A_F_Manual : ARRAY[0..10] OF Bool;  (* 手動【Y701】A(左側) 高さ検査押え行： *)
    Out_CYw_HgtInsp_Clp_A_F_Done : BOOL;  (* 【Y701】A(左側) 高さ検査押え行 動作完了 *)
    Out_CYw_HgtInsp_Lf_A_H_Auto : ARRAY[0..10] OF Bool;  (* 自動【Y702】A(左側) 高さ検査持上戻：; [1] 原点位置移動 *)
    Out_CYw_HgtInsp_Lf_A_H_Manual : ARRAY[0..10] OF Bool;  (* 手動【Y702】A(左側) 高さ検査持上戻： *)
    Out_CYw_HgtInsp_Lf_A_H_Done : BOOL;  (* 【Y702】A(左側) 高さ検査持上戻 動作完了 *)
    Out_CYw_HgtInsp_Lf_A_F_Auto : ARRAY[0..10] OF Bool;  (* 自動【Y703】A(左側) 高さ検査持上行：; [1] 高さ検査位置 *)
    Out_CYw_HgtInsp_Lf_A_F_Manual : ARRAY[0..10] OF Bool;  (* 手動【Y703】A(左側) 高さ検査持上行： *)
    Out_CYw_Sply_Slide_A_F_Auto : ARRAY[0..10] OF Bool;  (* 自動【Y617】A(左側) 供給スライド行：; [1] ワーク搬送 *)
    Out_CYw_Sply_Slide_A_F_Manual : ARRAY[0..10] OF Bool;  (* 手動【Y617】A(左側) 供給スライド行： *)
    Out_CYw_Sply_Pick_A_H_Auto : ARRAY[0..10] OF Bool;  (* 自動【Y618】A(左側) 供給ピックアップ戻：; [1] 原点位置移動; [2] ワーク回収; [3] ワーク設置完了後 *)
    Out_CYw_Sply_Pick_A_H_Manual : ARRAY[0..10] OF Bool;  (* 手動【Y618】A(左側) 供給ピックアップ戻： *)
    Out_CYw_Sply_Pick_A_H_Done : BOOL;  (* 【Y618】A(左側) 供給ピックアップ戻 動作完了 *)
    Out_CYw_Sply_Pick_A_F_Auto : ARRAY[0..10] OF Bool;  (* 自動【Y619】A(左側) 供給ピックアップ行：; [1] ワーク回収; [2] ワーク搬送 *)
    Out_CYw_Sply_Pick_A_F_Manual : ARRAY[0..10] OF Bool;  (* 自動【Y619】A(左側) 供給ピックアップ行： *)
    Out_CYw_Sply_Pick_A_F_Done : BOOL;  (* 【Y619】A(左側) 供給ピックアップ行 動作完了 *)
    Out_CYw_Sup_Chuck_A_Cl_H_Auto : ARRAY[0..10] OF Bool;  (* 自動【Y620】A(左側) 供給チャック閉 戻：; [1] 原点位置移動; [2] ワーク搬送 *)
    Out_CYw_Sup_Chuck_A_Cl_H_Manual : ARRAY[0..10] OF Bool;  (* 手動【Y620】A(左側) 供給チャック閉 戻： *)
    Out_CYw_Sup_Chuck_A_Cl_H_Done : BOOL;  (* 【Y620】A(左側) 供給チャック閉 戻 動作完了 *)
    Out_CYw_Sup_Chuck_A_Cl_F_Auto : ARRAY[0..10] OF Bool;  (* 自動【Y621】A(左側) 供給チャック開 行：; [1] ワーク回収 *)
    Out_CYw_Sup_Chuck_A_Cl_F_Manual : ARRAY[0..10] OF Bool;  (* 手動【Y621】A(左側) 供給チャック開 行： *)
    Out_CYw_Sup_Chuck_A_Cl_F_Done : BOOL;  (* 【Y621】A(左側) 供給チャック開 行 動作完了 *)
    Out_CYw_Sply_Slide_B_H_Auto : ARRAY[0..10] OF Bool;  (* 自動【Y622】B(右側) 供給スライド戻： *)
    Out_CYw_Sply_Slide_B_H_Manual : ARRAY[0..10] OF Bool;  (* 手動【Y622】B(右側) 供給スライド行： *)
    Out_CYw_Sply_Slide_B_Done : BOOL;  (* 【Y622】B(右側) 供給スライド戻 動作完了 *)
    Out_CYw_Sply_Slide_B_F_Auto : ARRAY[0..10] OF Bool;  (* 自動【Y623】B(右側) 供給スライド行： *)
    Out_CYw_Sply_Slide_B_F_Manual : ARRAY[0..10] OF Bool;  (* 手動【Y623】B(右側) 供給スライド行： *)
    Out_TDC_Stop : BOOL;  (* 【Y628】プレス上死点停止; at IOBus://unit#6/Output Bit 32 bits/Output Bit 28 *)
    TEST_M : ARRAY[0..99] OF Bool;  (* [1] 非常停止; [0] 自動運転ON *)
    ST0_Sup_Start : BOOL;  (* ST0_動作開始 *)
    Station_A_Data : ARRAY[0..8] OF sData;  (* A(左側)ステーションデータ *)
    Cv_A_Data : ARRAY[0..8] OF sData;  (* A(左側)コンベアデータ *)
    Station_B_Data : ARRAY[0..8] OF sData;  (* B(右側)ステーションデータ *)
    Cv_B_Data : ARRAY[0..8] OF sData;  (* B(右側)コンベアデータ *)
    ST0_A_Sup_End : BOOL;  (* ST0 A 動作完了 *)
    Ins_A_Cv_M : ARRAY[0..99] OF Bool;  (* [4] コンベア 動作開始; [5] ST1ワーク確認完了; [6] ST1ワーク不一致エラー; [7] ST2ワーク確認完了; [9] ST3ワーク確認完了; [11] ST4ワーク確認完了; [13] ST5ワーク確認完了; [15] ST6ワーク確認完了; [17] ST7ワーク確認完了; [8] ST2ワーク不一致エラー; [10] ST3ワーク不一致エラー; [12] ST4ワーク不一致エラー; [14] ST5ワーク不一致エラー; [16] ST6ワーク不一致エラー; [18] ST7ワーク不一致エラー; [3] STデータ移動完了; [1] 全ストッパー戻 動作開始; [2] 全ストッパ戻 確認完了 *)
    Ins_A_Cv_Error : BOOL;  (* 検査コンベア ワーク不一致エラー *)
    Ins_A_Next_Cycle : BOOL;  (* A(左側)検査次サイクル *)
    ST0_A_Sup_Busy : BOOL;  (* ST0 A 動作中 *)
    FH_New_Messages_Available : BOOL;
    FH_Sysmac_Error_Status : BYTE;
    FH_Line0_Command_Request : BOOL;
    FH_Line0_Trigger : BOOL;
    FH_Line0_Flow_Command_Request : BOOL;
    FH_Line0_Error_Clear : BOOL;
    FH_Line0_Result_Set_Request : BOOL;
    FH_Line0_Command_Code : DWORD;
    FH_Line0_Command_Parameter_0 : DINT;
    FH_Line0_Command_Parameter_1 : DINT;
    FH_Line0_Command_Parameter_2 : DINT;
    FH_Line0_Command_Parameter_3 : DINT;
    FH_Line0_Command_Completion : BOOL;
    FH_Line0_Busy : BOOL;
    FH_Line0_Trigger_Ready : BOOL;
    FH_Line0_Total_Judgment : BOOL;
    FH_Line0_Run_Mode : BOOL;
    FH_Line0_Trigger_Ack : BOOL;
    FH_Line0_Command_Ready : BOOL;
    FH_Line0_Shutter_Output : BOOL;
    FH_Line0_Flow_Command_Completion : BOOL;
    FH_Line0_Flow_Command_Busy : BOOL;
    FH_Line0_Flow_Command_Wait : BOOL;
    FH_Line0_Error_Status : BOOL;
    FH_Line0_Result_Notification : BOOL;
    FH_Line0_Command_Code_Echo_Back : DWORD;
    FH_Line0_Response_Code : DWORD;
    FH_Line0_Response_Data_0 : DINT;
    FH_Line0_Error_Code : DWORD;
    FH_Line0_DINT_Result_Data_0 : DINT;
    FH_Line0_DINT_Result_Data_1 : DINT;
    FH_Line0_DINT_Result_Data_2 : DINT;
    FH_Line0_DINT_Result_Data_3 : DINT;
    FH_Line0_DINT_Result_Data_4 : DINT;
    FH_Line0_DINT_Result_Data_5 : DINT;
    FH_Line0_DINT_Result_Data_6 : DINT;
    FH_Line0_DINT_Result_Data_7 : DINT;
    FH_Line1_Command_Request : BOOL;
    FH_Line1_Trigger : BOOL;
    FH_Line1_Flow_Command_Request : BOOL;
    FH_Line1_Error_Clear : BOOL;
    FH_Line1_Result_Set_Request : BOOL;
    FH_Line1_Command_Code : DWORD;
    FH_Line1_Command_Parameter_0 : DINT;
    FH_Line1_Command_Parameter_1 : DINT;
    FH_Line1_Command_Parameter_2 : DINT;
    FH_Line1_Command_Parameter_3 : DINT;
    FH_Line1_Command_Completion : BOOL;
    FH_Line1_Busy : BOOL;
    FH_Line1_Trigger_Ready : BOOL;
    FH_Line1_Total_Judgment : BOOL;
    FH_Line1_Run_Mode : BOOL;
    FH_Line1_Trigger_Ack : BOOL;
    FH_Line1_Command_Ready : BOOL;
    FH_Line1_Shutter_Output : BOOL;
    FH_Line1_Flow_Command_Completion : BOOL;
    FH_Line1_Flow_Command_Busy : BOOL;
    FH_Line1_Flow_Command_Wait : BOOL;
    FH_Line1_Error_Status : BOOL;
    FH_Line1_Result_Notification : BOOL;
    FH_Line1_Command_Code_Echo_Back : DWORD;
    FH_Line1_Response_Code : DWORD;
    FH_Line1_Response_Data_0 : DINT;
    FH_Line1_Error_Code : DWORD;
    FH_Line1_DINT_Result_Data_0 : DINT;
    FH_Line1_DINT_Result_Data_1 : DINT;
    FH_Line1_DINT_Result_Data_2 : DINT;
    FH_Line1_DINT_Result_Data_3 : DINT;
    FH_Line1_DINT_Result_Data_4 : DINT;
    FH_Line1_DINT_Result_Data_5 : DINT;
    FH_Line1_DINT_Result_Data_6 : DINT;
    FH_Line1_DINT_Result_Data_7 : DINT;
    FH_Line2_Command_Request : BOOL;
    FH_Line2_Trigger : BOOL;
    FH_Line2_Flow_Command_Request : BOOL;
    FH_Line2_Error_Clear : BOOL;
    FH_Line2_Result_Set_Request : BOOL;
    FH_Line2_Command_Code : DWORD;
    FH_Line2_Command_Parameter_0 : DINT;
    FH_Line2_Command_Parameter_1 : DINT;
    FH_Line2_Command_Parameter_2 : DINT;
    FH_Line2_Command_Parameter_3 : DINT;
    FH_Line2_Command_Completion : BOOL;
    FH_Line2_Busy : BOOL;
    FH_Line2_Trigger_Ready : BOOL;
    FH_Line2_Total_Judgment : BOOL;
    FH_Line2_Run_Mode : BOOL;
    FH_Line2_Trigger_Ack : BOOL;
    FH_Line2_Command_Ready : BOOL;
    FH_Line2_Shutter_Output : BOOL;
    FH_Line2_Flow_Command_Completion : BOOL;
    FH_Line2_Flow_Command_Busy : BOOL;
    FH_Line2_Flow_Command_Wait : BOOL;
    FH_Line2_Error_Status : BOOL;
    FH_Line2_Result_Notification : BOOL;
    FH_Line2_Command_Code_Echo_Back : DWORD;
    FH_Line2_Response_Code : DWORD;
    FH_Line2_Response_Data_0 : DINT;
    FH_Line2_Error_Code : DWORD;
    FH_Line2_DINT_Result_Data_0 : DINT;
    FH_Line2_DINT_Result_Data_1 : DINT;
    FH_Line2_DINT_Result_Data_2 : DINT;
    FH_Line2_DINT_Result_Data_3 : DINT;
    FH_Line2_DINT_Result_Data_4 : DINT;
    FH_Line2_DINT_Result_Data_5 : DINT;
    FH_Line2_DINT_Result_Data_6 : DINT;
    FH_Line2_DINT_Result_Data_7 : DINT;
    FH_Line3_Command_Request : BOOL;
    FH_Line3_Trigger : BOOL;
    FH_Line3_Flow_Command_Request : BOOL;
    FH_Line3_Error_Clear : BOOL;
    FH_Line3_Result_Set_Request : BOOL;
    FH_Line3_Command_Code : DWORD;
    FH_Line3_Command_Parameter_0 : DINT;
    FH_Line3_Command_Parameter_1 : DINT;
    FH_Line3_Command_Parameter_2 : DINT;
    FH_Line3_Command_Parameter_3 : DINT;
    FH_Line3_Command_Completion : BOOL;
    FH_Line3_Busy : BOOL;
    FH_Line3_Trigger_Ready : BOOL;
    FH_Line3_Total_Judgment : BOOL;
    FH_Line3_Run_Mode : BOOL;
    FH_Line3_Trigger_Ack : BOOL;
    FH_Line3_Command_Ready : BOOL;
    FH_Line3_Shutter_Output : BOOL;
    FH_Line3_Flow_Command_Completion : BOOL;
    FH_Line3_Flow_Command_Busy : BOOL;
    FH_Line3_Flow_Command_Wait : BOOL;
    FH_Line3_Error_Status : BOOL;
    FH_Line3_Result_Notification : BOOL;
    FH_Line3_Command_Code_Echo_Back : DWORD;
    FH_Line3_Response_Code : DWORD;
    FH_Line3_Response_Data_0 : DINT;
    FH_Line3_Error_Code : DWORD;
    FH_Line3_DINT_Result_Data_0 : DINT;
    FH_Line3_DINT_Result_Data_1 : DINT;
    FH_Line3_DINT_Result_Data_2 : DINT;
    FH_Line3_DINT_Result_Data_3 : DINT;
    FH_Line3_DINT_Result_Data_4 : DINT;
    FH_Line3_DINT_Result_Data_5 : DINT;
    FH_Line3_DINT_Result_Data_6 : DINT;
    FH_Line3_DINT_Result_Data_7 : DINT;
    FH_Line0_Command_Request_1 : BOOL;  (* A(左側) 出力：ST1 コマンド実行; at ECAT://node#4/Line0 Command Request *)
    FH_Line0_Trigger_1 : BOOL;  (* A(左側) 出力：ST1 測定トリガ; at ECAT://node#4/Line0 Trigger *)
    FH_Line0_Error_Clear_1 : BOOL;  (* A(左側) 出力：ST1 エラークリア; at ECAT://node#4/Line0 Error Clear *)
    FH_Line0_Command_Code_1 : DWORD;  (* 出力：コマンドコード; at ECAT://node#4/Line0 Command Code *)
    FH_Line0_Command_Completion_1 : BOOL;  (* A(左側) 入力：ST1 コマンド実行完了; at ECAT://node#4/Line0 Command Completion *)
    FH_Line0_Busy_1 : BOOL;  (* A(左側) 入力：ST1 処理実行中; at ECAT://node#4/Line0 Busy *)
    FH_Line0_Trigger_Ready_1 : BOOL;  (* A(左側) 入力：ST1 測定準備完了; at ECAT://node#4/Line0 Trigger Ready *)
    FH_Line0_Total_Judgment_1 : BOOL;  (* A(左側) 入力：ST1 総合判定; at ECAT://node#4/Line0 Total Judgment *)
    FH_Line0_Error_Status_1 : BOOL;  (* A(左側) 入力：ST1 エラー信号; at ECAT://node#4/Line0 Error Status *)
    FH_Line0_Result_Notification_1 : BOOL;  (* A(左側) 入力：ST1 出力完了; at ECAT://node#4/Line0 Result Notification *)
    FH_Line0_DINT_Result_Data_0_1 : DINT;  (* A(左側) 入力：ST1 判定0結果; at ECAT://node#4/Line0 DINT Result Data 0 *)
    FH_Line0_DINT_Result_Data_1_1 : DINT;  (* A(左側) 入力：ST1 判定1結果; at ECAT://node#4/Line0 DINT Result Data 1 *)
    FH_Line0_DINT_Result_Data_2_1 : DINT;  (* A(左側) 入力：ST1 判定2結果; at ECAT://node#4/Line0 DINT Result Data 2 *)
    FH_Line0_DINT_Result_Data_3_1 : DINT;  (* A(左側) 入力：ST1 判定3結果; at ECAT://node#4/Line0 DINT Result Data 3 *)
    FH_Line0_DINT_Result_Data_4_1 : DINT;  (* A(左側) 入力：ST1 判定4結果; at ECAT://node#4/Line0 DINT Result Data 4 *)
    FH_Line0_DINT_Result_Data_5_1 : DINT;  (* A(左側) 入力：ST1 判定5結果; at ECAT://node#4/Line0 DINT Result Data 5 *)
    FH_Line0_DINT_Result_Data_6_1 : DINT;  (* A(左側) 入力：ST1 判定6結果; at ECAT://node#4/Line0 DINT Result Data 6 *)
    FH_Line0_DINT_Result_Data_7_1 : DINT;  (* A(左側) 入力：ST1 判定7結果; at ECAT://node#4/Line0 DINT Result Data 7 *)
    FH_Line1_Command_Request_1 : BOOL;  (* A(左側) 出力：ST5 コマンド実行; at ECAT://node#4/Line1 Command Request *)
    FH_Line1_Trigger_1 : BOOL;  (* A(左側) 出力：ST5 測定トリガ; at ECAT://node#4/Line1 Trigger *)
    FH_Line1_Error_Clear_1 : BOOL;  (* A(左側) 出力：ST5 エラークリア; at ECAT://node#4/Line1 Error Clear *)
    FH_Line1_Command_Code_1 : DWORD;  (* at ECAT://node#4/Line1 Command Code *)
    FH_Line1_Command_Completion_1 : BOOL;  (* A(左側) 入力：ST5 コマンド実行完了; at ECAT://node#4/Line1 Command Completion *)
    FH_Line1_Busy_1 : BOOL;  (* A(左側) 入力：ST5 処理実行中; at ECAT://node#4/Line1 Busy *)
    FH_Line1_Trigger_Ready_1 : BOOL;  (* A(左側) 入力：ST5 測定準備完了; at ECAT://node#4/Line1 Trigger Ready *)
    FH_Line1_Total_Judgment_1 : BOOL;  (* A(左側) 入力：ST5 総合判定; at ECAT://node#4/Line1 Total Judgment *)
    FH_Line1_Error_Status_1 : BOOL;  (* A(左側) 入力：ST5 エラー信号; at ECAT://node#4/Line1 Error Status *)
    FH_Line1_Result_Notification_1 : BOOL;  (* A(左側) 入力：ST51 出力完了; at ECAT://node#4/Line1 Result Notification *)
    FH_Line1_DINT_Result_Data_0_1 : DINT;  (* A(左側) 入力：ST5 判定0結果; at ECAT://node#4/Line1 DINT Result Data 0 *)
    FH_Line1_DINT_Result_Data_1_1 : DINT;  (* A(左側) 入力：ST5 判定1結果; at ECAT://node#4/Line1 DINT Result Data 1 *)
    FH_Line1_DINT_Result_Data_2_1 : DINT;  (* A(左側) 入力：ST5 判定2結果; at ECAT://node#4/Line1 DINT Result Data 2 *)
    FH_Line1_DINT_Result_Data_3_1 : DINT;  (* A(左側) 入力：ST5 判定3結果; at ECAT://node#4/Line1 DINT Result Data 3 *)
    FH_Line1_DINT_Result_Data_4_1 : DINT;  (* A(左側) 入力：ST5 判定4結果; at ECAT://node#4/Line1 DINT Result Data 4 *)
    FH_Line1_DINT_Result_Data_5_1 : DINT;  (* A(左側) 入力：ST5 判定5結果; at ECAT://node#4/Line1 DINT Result Data 5 *)
    FH_Line1_DINT_Result_Data_6_1 : DINT;  (* A(左側) 入力：ST5 判定6結果; at ECAT://node#4/Line1 DINT Result Data 6 *)
    FH_Line1_DINT_Result_Data_7_1 : DINT;  (* A(左側) 入力：ST5 判定7結果; at ECAT://node#4/Line1 DINT Result Data 7 *)
    FH_Line2_Command_Request_1 : BOOL;  (* B(右側) 出力：ST1 コマンド実行; at ECAT://node#4/Line2 Command Request *)
    FH_Line2_Trigger_1 : BOOL;  (* B(右側) 出力：ST1 測定トリガ; at ECAT://node#4/Line2 Trigger *)
    FH_Line2_Error_Clear_1 : BOOL;  (* B(右側) 出力：ST1 エラークリア; at ECAT://node#4/Line2 Error Clear *)
    FH_Line2_Command_Completion_1 : BOOL;  (* B(右側) 入力：ST1 コマンド実行完了; at ECAT://node#4/Line2 Command Completion *)
    FH_Line2_Busy_1 : BOOL;  (* B(右側) 入力：ST1 処理実行中; at ECAT://node#4/Line2 Busy *)
    FH_Line2_Trigger_Ready_1 : BOOL;  (* B(右側) 入力：ST1 測定準備完了; at ECAT://node#4/Line2 Trigger Ready *)
    FH_Line2_Total_Judgment_1 : BOOL;  (* B(右側) 入力：ST1 総合判定; at ECAT://node#4/Line2 Total Judgment *)
    FH_Line2_Error_Status_1 : BOOL;  (* B(右側) 入力：ST1 エラー信号; at ECAT://node#4/Line2 Error Status *)
    FH_Line2_Result_Notification_1 : BOOL;  (* B(右側) 入力：ST1 出力完了; at ECAT://node#4/Line2 Result Notification *)
    FH_Line2_DINT_Result_Data_0_1 : DINT;  (* B(右側) 入力：ST1 判定0結果; at ECAT://node#4/Line2 DINT Result Data 0 *)
    FH_Line2_DINT_Result_Data_1_1 : DINT;  (* B(右側) 入力：ST1 判定1結果; at ECAT://node#4/Line2 DINT Result Data 1 *)
    FH_Line2_DINT_Result_Data_2_1 : DINT;  (* B(右側) 入力：ST1 判定2結果; at ECAT://node#4/Line2 DINT Result Data 2 *)
    FH_Line2_DINT_Result_Data_3_1 : DINT;  (* B(右側) 入力：ST1 判定3結果; at ECAT://node#4/Line2 DINT Result Data 3 *)
    FH_Line2_DINT_Result_Data_4_1 : DINT;  (* B(右側) 入力：ST1 判定4結果; at ECAT://node#4/Line2 DINT Result Data 4 *)
    FH_Line2_DINT_Result_Data_5_1 : DINT;  (* B(右側) 入力：ST1 判定5結果; at ECAT://node#4/Line2 DINT Result Data 5 *)
    FH_Line2_DINT_Result_Data_6_1 : DINT;  (* B(右側) 入力：ST1 判定6結果; at ECAT://node#4/Line2 DINT Result Data 6 *)
    FH_Line2_DINT_Result_Data_7_1 : DINT;  (* B(右側) 入力：ST1 判定7結果; at ECAT://node#4/Line2 DINT Result Data 7 *)
    FH_Line3_Command_Request_1 : BOOL;  (* B(右側) 出力：ST5 コマンド実行; at ECAT://node#4/Line3 Command Request *)
    FH_Line3_Trigger_1 : BOOL;  (* B(右側) 出力：ST5 測定トリガ; at ECAT://node#4/Line3 Trigger *)
    FH_Line3_Error_Clear_1 : BOOL;  (* B(右側) 出力：ST5 エラークリア; at ECAT://node#4/Line3 Error Clear *)
    FH_Line3_Command_Completion_1 : BOOL;  (* B(右側) 入力：ST5 コマンド実行完了; at ECAT://node#4/Line3 Command Completion *)
    FH_Line3_Busy_1 : BOOL;  (* B(右側) 入力：ST5 処理実行中; at ECAT://node#4/Line3 Busy *)
    FH_Line3_Trigger_Ready_1 : BOOL;  (* B(右側) 入力：ST5 測定準備完了; at ECAT://node#4/Line3 Trigger Ready *)
    FH_Line3_Total_Judgment_1 : BOOL;  (* B(右側) 入力：ST5 総合判定; at ECAT://node#4/Line3 Total Judgment *)
    FH_Line3_Error_Status_1 : BOOL;  (* B(右側) 入力：ST5 エラー信号; at ECAT://node#4/Line3 Error Status *)
    FH_Line3_Result_Notification_1 : BOOL;  (* B(右側) 入力：ST5 出力完了; at ECAT://node#4/Line3 Result Notification *)
    FH_Line3_DINT_Result_Data_0_1 : DINT;  (* B(右側) 入力：ST5 判定0結果; at ECAT://node#4/Line3 DINT Result Data 0 *)
    FH_Line3_DINT_Result_Data_1_1 : DINT;  (* B(右側) 入力：ST5 判定1結果; at ECAT://node#4/Line3 DINT Result Data 1 *)
    FH_Line3_DINT_Result_Data_2_1 : DINT;  (* B(右側) 入力：ST5 判定2結果; at ECAT://node#4/Line3 DINT Result Data 2 *)
    FH_Line3_DINT_Result_Data_3_1 : DINT;  (* B(右側) 入力：ST5 判定3結果; at ECAT://node#4/Line3 DINT Result Data 3 *)
    FH_Line3_DINT_Result_Data_4_1 : DINT;  (* B(右側) 入力：ST5 判定4結果; at ECAT://node#4/Line3 DINT Result Data 4 *)
    FH_Line3_DINT_Result_Data_5_1 : DINT;  (* B(右側) 入力：ST5 判定5結果; at ECAT://node#4/Line3 DINT Result Data 5 *)
    FH_Line3_DINT_Result_Data_6_1 : DINT;  (* B(右側) 入力：ST5 判定6結果; at ECAT://node#4/Line3 DINT Result Data 6 *)
    FH_Line3_DINT_Result_Data_7_1 : DINT;  (* B(右側) 入力：ST5 判定7結果; at ECAT://node#4/Line3 DINT Result Data 7 *)
    MdlChg : BOOL;  (* 機種切替：ON【GA120】 OFF【TE90】 *)
    FH_5552_10_A_Auto : BOOL;  (* ST1 FH測定開始 *)
    FH_A_ST1_Manual : BOOL;  (* ST1 *)
    FH_A_ST1_Done : BOOL;  (* ST1 画像検査完了 *)
    OriginDone : BOOL;  (* 原点復帰完了 *)
    DummyDone : BOOL;  (* ダミーチェック完了 *)
    HMI_CurrentPage : STRING[256];  (* HMI現在ページ *)
    Ins_A_End : BOOL;  (* A(左側)検査完了 *)
    Auto_A_Start : BOOL;  (* A(左側)自動運転 開始 *)
    Auto_Ready : BOOL;  (* 自動運転可能 *)
    ST1_A_Ca1_Busy : BOOL;  (* ST1 A検査中 *)
    ST1_A_Ca1_End : BOOL;  (* ST1 A 動作完了 *)
    ST2_A_Hgt_Busy : BOOL;  (* ST2 A 動作中 *)
    DLEP1_GT2_A_Auto : BOOL;
    DLEP1_IN : ARRAY[0..167] OF byte;  (* A(左側)GT2; [16] センサエラー; [48] 生データ; network input *)
    DLEP2_IN : ARRAY[0..167] OF byte;  (* B(右側)GT2; [16] センサエラー; [48] 生データ; network input *)
    DLEP1_OUT : ARRAY[0..79] OF BOOL;  (* A(左側)GT2; [0] ゼロリセット; [48] エラークリア; network output *)
    DLEP2_OUT : ARRAY[0..79] OF BOOL;  (* B(右側)GT2; [0] ゼロリセット; [48] エラークリア; network output *)
    DLEP2_IN_Error : BOOL;  (* B(右側)センサエラー *)
    DLEP1_IN_Error : BOOL;  (* A(右側)センサエラー *)
    GT2_A_CurrentVal : INT;  (* A(左側) 測定値 *)
    GT2_B_CurrentVal : INT;  (* B(右側) 測定値 *)
    Hgt_A_Ins_Data : LREAL;  (* A測定データに変換 *)
    Hgt_B_Ins_Data : LREAL;  (* B測定データに変換 *)
    Hgt_A_ComputedValueData : LREAL;  (* A測定データ+13.000mm 算定データ *)
    Hgt_B_ComputedValueData : LREAL;  (* B測定データ+13.000mm 算定データ *)
    Hight_LowerLimit : LREAL;  (* 高さ検査 下限値 *)
    Hight_UpperLimit : LREAL;  (* 高さ検査 上限値 *)
    TimerQ_In_Sen_Tray_Direction_Check : BOOL;  (* 【X1007】コンテナトレイ方向 *)
    ST2_A_Hgt_End : BOOL;  (* ST2 A 動作完了 *)
    ST3_A_Dis1_Busy : BOOL;  (* ST3 A 動作中 *)
    RC1_Receive_PDO_Mapping_ControlWord_6040_00 : UINT;
    RC1_Receive_PDO_Mapping_ControlWord_6040_00_1 : UINT;
    RC1_Receive_PDO_Mapping_Target_Position_607A_00 : DINT;  (* A(左側)NG1排出：目標位置 *)
    RC1_Receive_PDO_Mapping_Mode_of_operation_6060_00 : SINT;
    RC1_Receive_PDO_Mapping_Profile_velocity_6081_00 : UDINT;
    RC1_Receive_PDO_Mapping_Profile_acceleration_6083_00 : UDINT;
    RC1_Receive_PDO_Mapping_Profile_deceleration_6084_00 : UDINT;
    RC1_Receive_PDO_Mapping_Physical_outputs_60FE_01 : UDINT;
    RC1_Transmit_PDO_Mapping_StatusWord_6041_00 : UINT;
    RC1_Transmit_PDO_Mapping_Position_actual_value_6064_00 : DINT;
    RC1_Transmit_PDO_Mapping_Mode_of_operation_display_6061_00 : SINT;
    RC1_Transmit_PDO_Mapping_Following_error_actual_valu_60F4_00 : DINT;
    RC1_Transmit_PDO_Mapping_Torque_actual_value_6077_00 : INT;
    RC1_Transmit_PDO_Mapping_Digital_inputs_60FD_00 : UDINT;
    RC1_Transmit_PDO_Mapping_Error_code_603F_00 : UINT;
    RC2_Receive_PDO_Mapping_ControlWord_6040_00 : UINT;
    RC2_Receive_PDO_Mapping_Target_Position_607A_00 : DINT;
    RC2_Receive_PDO_Mapping_Mode_of_operation_6060_00 : SINT;
